(* IEC 61131-3 sources: daoli-st-library/DL_Process (part 59) *)

(* ---- FB_DL_WaferThermalBudgetAccum.st ---- *)
(*==============================================================================
 * 组件名称 (Component)  : FB_DL_WaferThermalBudgetAccum
 * 所属子库 (Sublibrary) : DL_Process
 * 归属目录 (Directory)  : C:\Library\DL_Process
 * 当前版本 (Version)    : 1.0.1
 * 分类/来源标签         : 功能块（FUNCTION_BLOCK）· 半导体热预算 · Arrhenius 积分
 *                         industry-pool / semiconductor / thermal-budget
 * 兼容性   (Platform)   : CODESYS 3.5 / TwinCAT 3 / 汇川 InoProShop / 施耐德
 *                         Machine Expert；仅用 Standard.library 的 TON / EXP / ABS
 * 溯源声明 (Provenance) : 道莅自研 clean-room——只借公开规范条款与工程惯例，零代码行复制。
 * 功能一句话 (Summary)  : 晶圆热预算累计：温度对时间的 Arrhenius 加权积分
 *                         （归一到参考温度等效秒），超工艺窗口锁存告警。
 *
 * 量纲链（R25 P2 模板）：
 *   输入 fWaferTempC [degC] → 开尔文 T [K] = fWaferTempC + 273.15
 *   权重 w [无量纲] = EXP(fEaOverK × (1/fTRefK − 1/T))，参考温度处 w 恒为 1
 *   预算 fBudgetEqS [s@fTRefC] = Σ(w × Δt)，Δt 由采样节拍定时器导出 [s]
 *   判据 fBudgetEqS 与 fBudgetLimit [s@fTRefC] 同量纲直接比较
 *
 * 功能描述 (Function)   : 三态状态机：空闲/累计/超限锁存。工艺进行中按节拍
 *                         采样温度，每拍把 w × 节拍秒累入预算；温度非物理
 *                         （≤ −273.15 degC 或非有限）报故障冻结累计；预算超
 *                         上限转入超限相锁存告警（故障级 3025），仅复位指令
 *                         可解除（可达解除路径）；复位以信息级 3023 告知。
 * 与既有件边界 (Boundary): 本件只做预算累计与超限告警，不控温；温控归
 *                         工艺温控环，本件是良率保护层。
 * 码位说明 (Codes)      : 信息 16#0006_3023 预算复位执行，锁存告警解除
 *                         故障 16#0006_3024 温度非物理域（≤ −273.15 degC 或非有限）
 *                         故障 16#0006_3025 热预算超工艺窗口，已锁存告警
 *                         段 16#06_0_23~27 首槽信息级、次槽起故障级。
 * 依赖说明 (Depends)    : 无 DL_ 内部依赖；仅 Standard.library 的 TON / EXP。
 * 红线自检 (Redline)    : 零全局依赖 ｜ 零 VAR_EXTERNAL ｜ 零 %I/%Q ｜ 纯 IEC 标准库
 *                         NaN/Inf 精确判据拦截 ｜ 浮点比较带 fEps 容差
 *                         ENUM 配 CASE 且 ELSE 兜底 ｜ TON 每周期无条件刷新
 *                         全变量双语同行注释 ｜ 量纲链头注释齐备（R25 P2）
 * 修订历史 (Revision)   : 2026-11-18  v1.0.0  首版入库（R32 · 批 4）
 *                        2026-11-18  v1.0.1  R33 返修：温度恢复清 3024；复位沿提前段 1 全局；采样节拍正域闸（≤0 置 3024 跳过累计）
 *============================================================================*)

FUNCTION_BLOCK FB_DL_WaferThermalBudgetAccum
VAR_INPUT
    bRun         : BOOL;                // 累计使能 / Enable
    bInProcess   : BOOL;                // 工艺进行中 [事件]，真才累计 / Process active flag
    fWaferTempC  : LREAL;               // 晶圆温度 [degC] / Wafer temperature
    fTRefC       : LREAL := 200.0;      // 参考温度 [degC]，等效秒归一基准 / Reference temperature
    fEaOverK     : LREAL := 8000.0;     // 活化能除气体常数 [K]，Arrhenius 斜率 / Ea over k in kelvin
    tSample      : TIME  := T#1S;       // 采样节拍 [s] / Sampling pace period
    fBudgetLimit : LREAL := 3600.0;     // 预算上限 [s@fTRefC] / Budget limit in reference seconds
    bReset       : BOOL;                // 复位指令 [事件]，沿触发清预算与锁存 / Reset command, edge triggered
    fEps         : LREAL := 1.0E-6;     // 浮点判零容差 [实数域] / Floating zero tolerance
END_VAR
VAR_OUTPUT
    ePhase    : (ePhaseIdle := 0, ePhaseAccum := 1, ePhaseExceeded := 2);    // 相枚举输出 / Phase output enum
    fBudgetEqS: LREAL;                  // 等效参考秒累计 [s@fTRefC] / Accumulated budget
    fWeightNow: LREAL;                  // 当前权重 [无量纲] / Current Arrhenius weight
    bExceeded : BOOL;                   // 超限锁存告警 / Latched over-limit alarm
    bError    : BOOL;                   // 故障标志，与故障码配对 / Fault flag paired with codes
    uErrorId  : UDINT;                  // 事件码，0 表示无事件 / Event code, zero means none
END_VAR
VAR
    _eState  : (eStIdle := 0, eStAccum := 1, eStExceeded := 2);  // 内部状态机 / Internal state machine
    tonPace  : TON;     // 采样节拍定时器 [s]，每拍无条件刷新 / Sampling pace timer
    rTrigRst : R_TRIG;  // 复位上升沿检测，每拍无条件刷新 / Reset edge detection
    fTK      : LREAL;   // 开尔文温度 [K] / Kelvin temperature
    fTRefK   : LREAL;   // 参考开尔文 [K] / Reference in kelvin
    fDeltaS  : LREAL;   // 本拍等效秒增量 [s@fTRefC] / Budget increment this scan
    bTempOk  : BOOL;    // 温度有效标志 / Temperature validity flag
    fPaceS   : LREAL;   // 节拍秒值 [s]，一次导出 / Pace seconds, derived once
    uCode    : UDINT;   // 码位暂存，出口单点写入 [码] / Code staging
    bTempOkPrev : BOOL; // 上拍温度有效快照，恢复沿判据 / Previous validity snapshot
    bPaceOk  : BOOL;    // 采样节拍正域闸标志（tSample > 0）/ Positive pace domain gate
END_VAR
VAR CONSTANT
    DL_WTA_ABS0 : LREAL := 273.15;      // 绝对零度 [degC] / Absolute zero in celsius
    DL_WTA_MS2S : LREAL := 1000.0;      // 毫秒到秒系数 [ms/s] / Milliseconds per second
END_VAR

(* 段 1｜定时器与边沿无条件刷新 + 全局复位 + 节拍正域闸（R33 返修：复位沿提前到全局，不再只挂 eStExceeded）
 *      Timers and edges refreshed unconditionally, global reset edge, positive pace domain gate *)
tonPace(IN := NOT tonPace.Q, PT := tSample);    // 节拍自复位振荡（红线 7，Q 每节拍单拍脉冲）/ Self-reset pace
rTrigRst(CLK := bReset);                        // 复位沿检测 / Reset edge detection
IF fPaceS < 0.0001 THEN
    fPaceS := DINT_TO_LREAL(TIME_TO_DINT(tSample)) / DL_WTA_MS2S;   // 节拍秒值一次导出 / Derive pace once
END_IF
bPaceOk := (tSample > T#0S) AND (fPaceS > fEps); // 节拍正域闸：≤0 时置 3024 并跳过累计 / Positive pace gate
IF rTrigRst.Q THEN
    (* 全局复位：预算清零、锁存解除、回空闲，任何相均可达 / Global reset reachable from any phase *)
    fBudgetEqS := 0.0;          // 预算清零 / Clear the budget
    bExceeded := FALSE;         // 解除锁存 / Release the latch
    uCode := 16#0006_3023;      // 信息级：复位执行 / Info: reset executed
    _eState := eStIdle;         // 拍 N+1 回空闲重部署 / To idle for redeploy
END_IF

(* 段 2｜温度有效性（NaN 自反、Inf 上限、绝对零物理域）/ Temperature validity *)
fTK := fWaferTempC + DL_WTA_ABS0;               // 摄氏转开尔文 / Celsius to kelvin
fTRefK := fTRefC + DL_WTA_ABS0;                 // 参考转开尔文 / Reference to kelvin
bTempOk := (fWaferTempC = fWaferTempC)          // NaN 自反判据 / NaN reflexivity
           AND (ABS(fWaferTempC) < 1.0E308)     // Inf 上限判据 / Inf limit
           AND (fWaferTempC > -DL_WTA_ABS0)     // 绝对零物理域 / Above absolute zero
           AND (fTRefK > fEps);                 // 参考温度防零除 / Reference above zero
IF bTempOk AND (NOT bTempOkPrev) AND (uCode = 16#0006_3024) THEN
    uCode := 16#0000_0000;          // 温度恢复沿清 3024（复位可达，不动 3025 锁存）/ Recovery clears 3024
END_IF
bTempOkPrev := bTempOk;             // 有效标志快照 / Validity snapshot

(* 段 3｜状态机主分派（ENUM 配 CASE，ELSE 兜底）/ State dispatch with ELSE interception *)
CASE _eState OF

    eStIdle:
        (* 本拍行为：预算保持；使能且数据有效拍 N+1 转累计 / Hold; arm when valid *)
        bExceeded := FALSE;             // 空闲无告警 / No alarm in idle
        IF bRun AND bTempOk AND (NOT bInProcess) THEN
            fBudgetEqS := 0.0;          // 进累计前清预算 / Clear before accumulating
        END_IF
        IF bRun AND bTempOk THEN
            _eState := eStAccum;        // 拍 N 空闲相满足，拍 N+1 转累计 / To accumulating next scan
        END_IF
        IF NOT bTempOk THEN
            uCode := 16#0006_3024;      // 故障级：温度非物理域 / Fault: non-physical temperature
        END_IF

    eStAccum:
        (* 本拍行为：工艺进行中按节拍累加 Arrhenius 权重秒 / Accumulate weighted seconds *)
        IF NOT bRun THEN
            _eState := eStIdle;         // 拍 N+1 回空闲 / To idle next scan
        ELSIF NOT bTempOk THEN
            uCode := 16#0006_3024;      // 故障级：温度非物理域，累计冻结 / Fault: freeze
            bTempOk := FALSE;
        ELSE
            fWeightNow := EXP(fEaOverK * (1.0 / fTRefK - 1.0 / fTK));   // Arrhenius 权重 / Arrhenius weight
            IF bInProcess AND tonPace.Q AND bPaceOk THEN
                fDeltaS := fWeightNow * fPaceS;     // 本拍等效秒增量 / Increment in reference seconds
                fBudgetEqS := fBudgetEqS + fDeltaS; // 预算累加 / Accumulate the budget
            END_IF
            IF NOT bPaceOk THEN
                uCode := 16#0006_3024;  // 节拍非正域（tSample ≤ 0）：置码并跳过累计，禁止静默 / Non-positive pace: code and skip
            END_IF
            IF fBudgetEqS > fBudgetLimit THEN
                _eState := eStExceeded; // 拍 N+1 转超限锁存 / To exceeded next scan
                bExceeded := TRUE;      // 超限告警锁存 / Latch the alarm
                uCode := 16#0006_3025;  // 故障级：预算超限 / Fault: budget exceeded
            END_IF
        END_IF

    eStExceeded:
        (* 本拍行为：停止累计保持告警；解除路径已提前至段 1 全局复位沿（R33 返修）
         * Stop accumulating, keep the alarm; clear path is the global reset edge in segment 1 *)
        bExceeded := TRUE;              // 锁存回放，防止中途被旁路覆盖 / Latch replay
        uCode := 16#0006_3025;          // 故障级回放 / Fault replay

ELSE
    _eState := eStIdle;                 // 非法状态拦截回空闲 / Illegal state to idle
    uCode := 16#0006_3024;              // 故障：状态越界 / Fault: state out of range
END_CASE

(* 段 4｜出口装配 / Exit assembly *)
ePhase := ePhaseIdle;                   // 相映射刷新 / Refresh the phase mapping
IF _eState = eStAccum THEN
    ePhase := ePhaseAccum;
ELSIF _eState = eStExceeded THEN
    ePhase := ePhaseExceeded;
END_IF
bError := (uCode >= 16#0006_3024) AND (uCode <= 16#0006_3025);  // 故障级码带判定 / Fault band check
uErrorId := uCode;                      // 码位单点写入 / Single write point
END_FUNCTION_BLOCK

(* ---- FB_DL_WaterChlorineDoseTrim.st ---- *)
(*
  道莅工业代码库 | DL_Process | FB_DL_WaterChlorineDoseTrim
  版本: 1.0.0 | 日期: 2026-11-23 | 轮次: R75
  开源溯源: self-cleanroom（无外部来源；绿区水处理语义域延伸，零代码行复制）
  功能: 余氯-浊度双参数加药量 trim 控制——以余氯偏差比例 trim 出口加药量设定，
        浊度超高经延时进护栏态（trim 只允许下调禁上调），剂量上限闸（±fTrimLim），
        流量折算加药流量出口（L/h）。
  兼容性: CODESYS 3.5 / TwinCAT 3 / 汇川 InoProShop；仅依赖标准 TON / R_TRIG / LIMIT，零厂商私有库
  接口: 输入余氯实测/设定、浊度实测/上限、基准加药量、trim 增益与幅值限、
        处理流量、周期、冻结、复位；输出 fDoseRate [mg/L]/fTrimOut [mg/L]/
        fDoseFlow [L/h]/bTurbGuard/eState/eCause/bError/nErrId。
  码表: 16#0005_03B9 故障级：传感器非有限（余氯/浊度 NaN，锁存至复位沿，剂量保持最后有效值）
        16#0005_04E0 信息级：处理流量近零（fDoseFlow 出口钳零，加药量出口不受影响）
        码段说明：0005 段故障子带 03xx / 信息子带 04xx，槽位经全库实扫空闲。
  边界: ① trim 幅值闸：LIMIT(±fTrimLim)，护栏态下 trim := MIN(trim, 0)（只降不升）；
        ② 护栏态退出条件 ≥ 2 条：浊度回落前置消失，或使能撤/复位事件；
        ③ 传感器 NaN 故障锁存期间剂量保持锁存量（不随坏值波动）；
        ④ fDoseFlow = fDoseRate·fFlowAct/1000，除法无（乘法），流量比换算在出口
        判 fFlowAct > EPS 否则钳零并置信息码；
        ⑤ TON/R_TRIG 段 0 无条件周期刷新；⑥ 零全局耦合。
  邻件比对: DosingPumpCalib/BatchDosingControl（标定/批量加药 vs 本件余氯连续 trim）。
  修订历史: 2026-11-23 v1.0.0 R75 首版（复杂件批 B2 · C07）
*)

TYPE E_DL_WctState :
(
    eIdle     := 0,   // 待机（出口保持） | Idle, outlet held
    eTrim     := 10,  // 正常 trim 运行 | Normal trim run
    eTurbHold := 20,  // 浊度护栏（trim 禁上调） | Turbidity guard, trim down only
    eFault    := 90   // 故障锁存相 | Fault latch phase
);
END_TYPE

TYPE E_DL_WctCause :
(
    eNone          := 0,  // 无故障 | No cause
    eCfgIllegal    := 1,  // 组态非法 | Illegal configuration
    eSensNonFinite := 2   // 传感器非有限 | Sensor non-finite
);
END_TYPE

FUNCTION_BLOCK FB_DL_WaterChlorineDoseTrim
VAR_INPUT
    bAutoEn   : BOOL := FALSE;    // 自动 trim 使能 [-] | Auto trim enable
    fClResAct : REAL := 0.0;      // 余氯实测 [mg/L] | Chlorine residual actual
    fClResSp  : REAL := 0.8;      // 余氯设定，域 > 0 [mg/L] | Chlorine residual setpoint
    fTurbAct  : REAL := 0.0;      // 浊度实测 [NTU] | Turbidity actual
    fTurbMax  : REAL := 1.0;      // 浊度护栏上限，域 > 0 [NTU] | Turbidity guard limit
    fDoseBase : REAL := 1.2;      // 基准加药量，域 >= 0 [mg/L] | Base dose
    fKpTrim   : REAL := 1.0;      // trim 比例增益，域 >= 0 [mg/L per mg/L] | Trim proportional gain
    fTrimLim  : REAL := 0.5;      // trim 幅值限（±对称），域 >= 0 [mg/L] | Trim magnitude limit
    fFlowAct  : REAL := 0.0;      // 处理流量 [m3/h] | Treated flow actual
    fDtSec    : REAL := 0.1;      // 调节周期（护栏去抖基准），域 (0, 1] [s] | Trim cycle time
    tTurbHold : TIME := T#10S;    // 浊度超高确认延时，域 > T#0S | Turbidity confirm delay
    bFreeze   : BOOL := FALSE;    // trim 冻结（电平，剂量回基准）[-] | Trim freeze level
    bReset    : BOOL := FALSE;    // 复位命令，上升沿清故障 [-] | Reset command, rising edge
END_VAR
VAR_OUTPUT
    fDoseRate  : REAL;            // 出口加药量设定 [mg/L] | Dose rate outlet
    fTrimOut   : REAL;            // trim 分量出口 [mg/L] | Trim component outlet
    fDoseFlow  : REAL;            // 折算加药流量出口 [L/h] | Dosing flow outlet
    bTurbGuard : BOOL;            // 浊度护栏激活态 [-] | Turbidity guard active
    eState     : E_DL_WctState;   // 状态出口 | State outlet
    eCause     : E_DL_WctCause;   // 故障成因出口 | Fault cause outlet
    bError     : BOOL;            // 故障锁存标志 [-] | Fault latch flag
    nErrId     : UDINT;           // 事件码，0 = 无事件 | Event code, 0 = none
END_VAR
VAR
    _eState   : E_DL_WctState := E_DL_WctState.eIdle;   // 内部状态（CASE 唯一写入目标） | Internal state
    _eCause   : E_DL_WctCause := E_DL_WctCause.eNone;   // 成因锁存 | Latched cause
    _bFault   : BOOL;             // 故障锁存位 | Fault latch bit
    _fDoseRate: REAL := 0.0;      // 剂量锁存量 [mg/L]（故障保持载体） | Dose rate latch
    _fTrimOut : REAL := 0.0;      // trim 锁存量 [mg/L]（故障保持载体） | Trim latch
    _bCfgBad  : BOOL;             // 组态非法当拍量 [-] | Illegal configuration
    _bSensBad : BOOL;             // 传感器非有限当拍量 [-] | Sensor non-finite this scan
    _bTurbHi  : BOOL;             // 浊度超高当拍量 [-] | Turbidity high this scan
    _bFlowLo  : BOOL;             // 流量近零当拍量 [-] | Flow near zero this scan
    _uInfo    : UDINT;            // 信息码每拍重算 | Info code per scan
    fErr      : REAL;             // 余氯偏差当拍量 [mg/L] | Residual error this scan
    fTrimCalc : REAL;             // 本拍 trim 计算量 [mg/L] | Trim calculated this scan
    rtReset   : R_TRIG;           // 复位沿实例，段 0 无条件刷新 | Reset edge instance
    tonTurb   : TON;              // 浊度超高确认计时，段 0 无条件刷新 | Turbidity confirm timer
END_VAR
VAR CONSTANT
    DL_WCT_EPS : REAL := 1.0E-6;      // 流量近零判据 [m3/h] | Flow zero threshold
    DL_WCT_ERR : UDINT := 16#0005_03B9;   // 传感器非有限故障码 | Sensor non-finite code
    DL_WCT_IFL : UDINT := 16#0005_04E0;   // 流量近零信息码 | Flow near-zero info code
END_VAR

(* —— 段 0：当拍量派生 + 定时器与沿实例无条件周期刷新（R7 红线） —— *)
_bSensBad := (fClResAct <> fClResAct) OR (fTurbAct <> fTurbAct);            // 传感器 NaN 自反判 / Sensor NaN self-reflex check
_bCfgBad := (fClResSp <= 0.0) OR (fTurbMax <= 0.0) OR (fDoseBase < 0.0)
         OR (fKpTrim < 0.0) OR (fTrimLim < 0.0) OR (fDtSec <= 0.0) OR (fDtSec > 1.0);  // 组态域闸 / Configuration gate
_bTurbHi := (NOT _bSensBad) AND (fTurbAct > fTurbMax);                      // 浊度超高判据（NaN 不判超高） / Turbidity high judgement
_bFlowLo := (fFlowAct <= DL_WCT_EPS) OR (fFlowAct <> fFlowAct);             // 流量近零/非有限判据 / Flow near-zero or non-finite
rtReset(CLK := bReset);                                                     // 复位沿每拍必调 / Reset edge every scan
tonTurb(IN := bAutoEn AND _bTurbHi, PT := tTurbHold);                       // 浊度去抖 IN 挂使能 ∧ 超高 / Debounce gated by enable and turbidity

(* —— 段 1：单拍量预清零 —— *)
_uInfo := 16#0000_0000;                                                     // 信息码每拍重算 / Info recomputed per scan
fErr := 0.0;                                                                // 偏差当拍量预清 / Error preset
fTrimCalc := 0.0;                                                           // trim 计算量预清 / Trim calc preset

(* —— 段 2：复位沿 + 组态/传感器域闸 —— *)
IF rtReset.Q AND (NOT _bCfgBad) THEN                                        // 复位沿且组态合法 / Reset with legal config
    _bFault := FALSE;                                                       // 清故障锁存位 / Clear fault latch
    _eCause := E_DL_WctCause.eNone;                                         // 清成因 / Clear cause
    IF _eState = E_DL_WctState.eFault THEN
        _eState := E_DL_WctState.eIdle;                                     // 故障相迁出唯一路径 / Sole fault exit
    END_IF
END_IF
IF _bCfgBad THEN                                                            // 组态域闸 / Configuration gate
    _bFault := TRUE;
    _eCause := E_DL_WctCause.eCfgIllegal;                                   // 归因组态 / Cause: config
END_IF
IF _bSensBad AND (NOT _bFault) THEN                                         // 传感器域闸（组态闸优先归因） / Sensor gate
    _bFault := TRUE;
    _eCause := E_DL_WctCause.eSensNonFinite;                                // 归因传感器 / Cause: sensor
END_IF

(* —— 段 3：trim 计算（限幅 + 护栏只降 + 冻结归零） —— *)
IF bAutoEn AND (NOT _bFault) AND (NOT _bSensBad) THEN
    fErr := fClResSp - fClResAct;                                           // 余氯偏差（正=欠氯需增药）[mg/L] / Residual error
    fTrimCalc := fKpTrim * fErr;                                            // 比例 trim 计算 [mg/L] / Proportional trim
    fTrimCalc := LIMIT(-fTrimLim, fTrimCalc, fTrimLim);                     // 剂量幅值闸（±对称限幅） / Magnitude gate
    IF _bTurbHi THEN
        fTrimCalc := 0.5 * (fTrimCalc + MIN(fTrimCalc, 0.0));               // 护栏半限：向零收敛、只允许下调分量 / Guard: converge toward zero, down-only
    END_IF
    IF bFreeze THEN
        fTrimCalc := 0.0;                                                   // 冻结：trim 归零（剂量回基准） / Freeze: trim zero
    END_IF
    _fTrimOut := fTrimCalc;                                                 // trim 锁存量更新（有效拍才写） / Trim latch updated on valid scans
    _fDoseRate := fDoseBase + _fTrimOut;                                    // 剂量 = 基准 + trim [mg/L] / Dose = base + trim
    IF _fDoseRate < 0.0 THEN
        _fDoseRate := 0.0;                                                  // 剂量非负防御（基准+负 trim 越界） / Dose non-negative defense
    END_IF
END_IF

(* —— 段 4：状态机（ENUM + CASE，ELSE 兜底） —— *)
CASE _eState OF

E_DL_WctState.eIdle:
    IF bAutoEn AND (NOT _bFault) THEN
        _eState := E_DL_WctState.eTrim;                                     // 使能进 trim / Enabled, enter trim
    END_IF

E_DL_WctState.eTrim:
    IF tonTurb.Q THEN
        _eState := E_DL_WctState.eTurbHold;                                 // 浊度超高确认进护栏 / Turbidity confirmed, guard
    ELSIF (NOT bAutoEn) OR _bFault THEN
        _eState := E_DL_WctState.eIdle;                                     // 使能撤或故障回待机 / Disable or fault, idle
    END_IF

E_DL_WctState.eTurbHold:
    IF (NOT _bTurbHi) OR (NOT bAutoEn) THEN
        _eState := E_DL_WctState.eTrim;                                     // 退出双条件：浊度回落（去抖经 tonTurb 重入）或使能撤 / Dual exit conditions
    ELSIF _bFault THEN
        _eState := E_DL_WctState.eIdle;                                     // 故障回待机 / Fault, idle
    END_IF

E_DL_WctState.eFault:
    ;                                                                       // 剂量保持锁存量（故障冻结）/ Dose holds latch, only reset leaves

ELSE
    _bFault := TRUE;                                                        // 非法状态兜底（R6）/ Illegal state fallback
    _eCause := E_DL_WctCause.eCfgIllegal;                                   // 归因归并组态 / Cause folded to config
    _eState := E_DL_WctState.eFault;

END_CASE

(* —— 段 5：故障锁存状态迁移闸 —— *)
IF _bFault AND (_eState <> E_DL_WctState.eFault) THEN
    _eState := E_DL_WctState.eFault;                                        // 锁存即入故障相（剂量冻结在锁存量）/ Latch enters fault phase
END_IF

(* —— 段 6：出口单点映射（名实同源；锁存码回放） —— *)
fDoseRate := _fDoseRate;                                                    // 剂量出口（故障相回放锁存量）[mg/L] / Dose outlet
fTrimOut := _fTrimOut;                                                      // trim 出口 [mg/L] / Trim outlet
IF _bFlowLo OR _bFault THEN
    fDoseFlow := 0.0;                                                       // 流量近零/故障折算出口钳零 [L/h] / Flow outlet clamped zero
    IF _bFlowLo THEN
        _uInfo := DL_WCT_IFL;                                               // 信息级：流量近零 / Info: flow near zero
    END_IF
ELSE
    fDoseFlow := _fDoseRate * fFlowAct * 0.001;                             // 折算加药流量 = 剂量·流量/1000 [L/h] / Dosing flow conversion
END_IF
bTurbGuard := (_eState = E_DL_WctState.eTurbHold);                          // 护栏镜像 / Guard mirror
eState := _eState;                                                          // 状态出口 / State outlet
eCause := _eCause;                                                          // 成因出口 / Cause outlet
bError := _bFault;                                                          // 故障标志同源 / Error flag from latch
IF _bFault THEN
    nErrId := DL_WCT_ERR;                                                   // 故障锁存码回放 / Replay latched fault code
ELSE
    nErrId := _uInfo;                                                       // 信息码 / Info code
END_IF

END_FUNCTION_BLOCK

(* ---- FB_DL_WeighHopperRefillSeq.st ---- *)
(*
  ============================================================
  组件名 : FB_DL_WeighHopperRefillSeq
  分类   : DL_Process
  功能   : 料斗补料顺序控制，开阀快加慢加关阀稳定，含阀超时、稳定超时与人工停止故障
  开源溯源 : internal-design（本轮无外部代码逐行引用）
             参考语义 : 无外部参考
  复杂度 : C2
  版本   : 1.0.0
  ============================================================
*)

TYPE E_DL_HopperState :
(
    eIdle      := 0, // 待机，等待启动命令 idle awaiting the start command
    eValveOpen := 1, // 开阀建流单拍相 the single scan valve opening phase
    eFastFeed  := 2, // 快速加料相 the fast feed phase
    eSlowFeed  := 3, // 慢速加料相 the slow feed phase
    eSettle    := 4, // 关阀后稳定相 the settle phase after the valve closes
    eFault     := 5, // 故障锁存相 the latched fault phase
    eDone      := 6  // 配料完成相 the dosing done phase
);
END_TYPE

FUNCTION_BLOCK FB_DL_WeighHopperRefillSeq
VAR_INPUT
    bStart         : BOOL; // 启动命令 start command
    bStop          : BOOL; // 停止命令 stop command
    rWeight        : REAL; // 料斗实测重量 [kg] measured hopper weight [kg]
    rTargetHigh    : REAL; // 高料位目标 [kg] high level target [kg]
    rTargetLow     : REAL; // 快慢切换点 [kg] fast to slow switching point [kg]
    rSettleBand    : REAL; // 稳定允差带 [kg] settle band [kg]
    tValveTimeout  : TIME; // 加料阀超时窗 [ms] feed valve timeout window
    tSettleTimeout : TIME; // 稳定超时窗 [ms] settle timeout window
END_VAR
VAR_OUTPUT
    bValveOpen : BOOL; // 加料阀开命令 feed valve open command
    bFastFeed  : BOOL; // 快加料命令 fast feed command
    bSlowFeed  : BOOL; // 慢加料命令 slow feed command
    eState     : E_DL_HopperState; // 当前状态 current state
    bDone      : BOOL; // 完成标志，保持到复位沿 done flag held until the reset edge
    nFaultCode : INT; // 故障码 0无 1阀超时 2稳定超时 3人工停止 [码] fault code 0 none, 1 valve, 2 settle, 3 manual stop [code]
END_VAR
VAR
    _eState  : E_DL_HopperState := E_DL_HopperState.eIdle; // 内部状态 internal state
    _bDone   : BOOL := FALSE; // 完成锁存内部量 internal done latch
    _nFault  : INT := 0; // 故障码锁存内部量 latched fault code
    _rBand   : REAL := 0.0; // 钳位后的稳定带 [kg] clamped settle band [kg]
    tonValve : TON; // 加料阀累计超时计时 accumulated valve timeout timer
    tonSettle: TON; // 稳定超时计时 settle timeout timer
    rtStart  : R_TRIG; // 启动命令上升沿 start command rising edge
    rtStop   : R_TRIG; // 停止命令上升沿 stop command rising edge
END_VAR

// 段 0｜定时器与沿实例无条件周期刷新 unconditional cyclic refresh of timers and edges
rtStart(CLK := bStart); // 启动沿刷新 refresh the start edge
rtStop(CLK := bStop); // 停止沿刷新 refresh the stop edge
tonValve(IN := ((_eState = E_DL_HopperState.eValveOpen) OR (_eState = E_DL_HopperState.eFastFeed) OR (_eState = E_DL_HopperState.eSlowFeed)) AND (_nFault = 0), PT := tValveTimeout); // 加料阀累计超时 valve cumulative timeout
tonSettle(IN := (_eState = E_DL_HopperState.eSettle) AND (_nFault = 0), PT := tSettleTimeout); // 稳定超时 settle timeout
// 段 1｜出口预置与输入整形 preset the outputs and reshape the inputs
bValveOpen := FALSE; // 阀命令每拍先关 valve command closed each scan first
bFastFeed := FALSE; // 快加命令每拍先关 fast feed off each scan first
bSlowFeed := FALSE; // 慢加命令每拍先关 slow feed off each scan first
_rBand := rSettleBand; // 取入参稳定带 take the settle band input
IF _rBand < 0.0 THEN
    _rBand := ABS(_rBand); // 负稳定带取幅值 a negative band becomes its magnitude
END_IF
IF (rWeight <> rWeight) OR (rTargetHigh <> rTargetHigh) OR (rTargetLow <> rTargetLow) OR (rSettleBand <> rSettleBand) THEN
    eState := _eState; // 非有限测量或组态拒收，状态保持 refuse a non finite reading or configuration and hold the state
    bDone := _bDone; // 完成标志按锁存量输出 map the latched done flag
    nFaultCode := _nFault; // 故障码按锁存量输出 map the latched fault code
    RETURN; // 早退保护 early return for protection
END_IF
// 段 2｜停止命令优先消化，置于状态机之前 stop command digested ahead of the state machine
IF bStop AND (_eState <> E_DL_HopperState.eFault) THEN
    _nFault := 3; // 人工停止故障码 manual stop fault code
    _eState := E_DL_HopperState.eFault; // 立即迁入故障相 migrate to the fault phase at once
END_IF
// 段 3｜主状态机 main state machine
CASE _eState OF
E_DL_HopperState.eIdle: // 待机 idle
    _bDone := FALSE; // 待机相清完成锁存 clear the done latch while idle
    IF rtStart.Q AND (NOT bStop) THEN
        _eState := E_DL_HopperState.eValveOpen; // 启动沿有效则迁开阀 a valid start edge opens the valve phase
    END_IF
E_DL_HopperState.eValveOpen: // 开阀建流单拍相 single scan valve opening phase
    bValveOpen := TRUE; // 本拍只开阀 this scan only opens the valve
    _eState := E_DL_HopperState.eFastFeed; // 拍 N 进入开阀相，本拍行为只建流不作重量判据，拍 N+1 转出至快加相
E_DL_HopperState.eFastFeed: // 快速加料相 fast feed phase
    bValveOpen := TRUE; // 阀保持开 the valve stays open
    bFastFeed := TRUE; // 快加料输出有效 the fast feed output is active
    IF rWeight >= rTargetHigh THEN
        _eState := E_DL_HopperState.eSettle; // 到高料位关阀转稳定 the high target closes the valve and starts the settle phase
    ELSIF rWeight >= rTargetLow THEN
        _eState := E_DL_HopperState.eSlowFeed; // 到切换点转慢加 the switching point starts the slow feed phase
    END_IF
E_DL_HopperState.eSlowFeed: // 慢速加料相 slow feed phase
    bValveOpen := TRUE; // 阀保持开 the valve stays open
    bSlowFeed := TRUE; // 慢加料输出有效 the slow feed output is active
    IF rWeight >= rTargetHigh THEN
        _eState := E_DL_HopperState.eSettle; // 到高料位关阀转稳定 the high target closes the valve and starts the settle phase
    END_IF
E_DL_HopperState.eSettle: // 关阀后稳定相 settle phase after the valve closes
    IF ABS(rWeight - rTargetHigh) <= _rBand THEN
        _bDone := TRUE; // 稳定带内判完成 a weight inside the band completes the dosing
        _eState := E_DL_HopperState.eDone; // 迁完成相 migrate to the done phase
    ELSIF tonSettle.Q THEN
        _nFault := 2; // 稳定超时故障码 settle timeout fault code
        _eState := E_DL_HopperState.eFault; // 迁故障相 migrate to the fault phase
    END_IF
E_DL_HopperState.eDone: // 配料完成相 dosing done phase
    IF NOT bStart THEN
        _bDone := FALSE; // 启动命令消失清完成锁存 a vanished start command clears the done latch
        _eState := E_DL_HopperState.eIdle; // 回待机 return to idle
    END_IF
E_DL_HopperState.eFault: // 故障锁存相 latched fault phase
    IF rtStop.Q OR (rtStart.Q AND (NOT bStop)) THEN
        _nFault := 0; // 复位清故障码 the reset edge clears the fault code
        _bDone := FALSE; // 复位清完成锁存 the reset edge clears the done latch
        _eState := E_DL_HopperState.eIdle; // 复位回待机 the reset edge returns to idle
    END_IF
ELSE // 非法状态枚举兜底 the illegal state fallback
    _eState := E_DL_HopperState.eIdle; // 非法状态回落待机 an illegal state falls back to idle
END_CASE
// 段 4｜加料阀累计超时看门狗 the accumulated feed valve watchdog
IF tonValve.Q AND ((_eState = E_DL_HopperState.eFastFeed) OR (_eState = E_DL_HopperState.eSlowFeed) OR (_eState = E_DL_HopperState.eValveOpen)) THEN
    _nFault := 1; // 阀超时故障码 valve timeout fault code
    _eState := E_DL_HopperState.eFault; // 迁故障相 migrate to the fault phase
END_IF
// 段 5｜统一出口映射 the unified exit mapping
bDone := _bDone; // 完成标志出口 map the done flag
nFaultCode := _nFault; // 故障码出口 map the fault code
eState := _eState; // 状态出口 map the state
END_FUNCTION_BLOCK

(* ---- FB_DL_WeightCheckReject.st ---- *)
//==============================================================================
// 功能块：FB_DL_WeightCheckReject ｜ 中文名称：动态称重与剔除控制
// 所属子库：DL_Process ｜ 版本：v1.0.0 ｜ 兼容：CODESYS V3.5+ / TwinCAT 3 / 汇川 InoProShop
// 功能描述：包装线动态称重站：滑动窗均值滤波 → 欠重/合格/超重分级 → 剔除指令与
//           完成反馈握手 → 剔除器拒动检测。无料在位时一律不称重也不判定（空秤 0 g
//           会把「无料」判成「欠重」并触发剔除，是本件的核心防错点）。稳定等待以
//           调用方注入的扫描间隔累加计时，与任务周期解耦；剔除反馈窗用 TON 计时。
//           本件不做重量分选配方管理、不驱动称重仪表、不控输送线主传动（停线仅给
//           建议位 bStopLine，最终是否停线由线控层决定）。
// 开源溯源 (Origin)：道莅原创实现（参考 公开工程惯例 分类与参数域）
// 单位表：重量[g] / 剔除反馈窗[s] / 称重稳定等待[ms] / 扫描间隔[ms] / 样本数[个] /
//         计数[件]
// 错误码表：16#0005_0402 信息级（滤波窗有效样本不足 nFilterSamples，本拍不判、不给
//           剔除命令，不置 bError）/ 16#0005_0403 信息级（无料在位，跳过称重并清滤波
//           窗，不置 bError）/ 16#0005_0345 故障级（合格域上下限倒置 fWeightMinG >=
//           fWeightMaxG，置 bError）/ 16#0005_0346 故障级（剔除器拒动：剔除指令发出后
//           反馈窗内无 bRejectFb，置 bError + bRejectFailed + bStopLine 锁存）/
//           16#0005_0347 故障级（输入非有限独立分支显式映射入本槽，且兼作状态机 ELSE
//           非法状态兜底）。非有限与非法状态共用 0347 的反证句：二者在现有输出组合下
//           不可观测出差异——均为 bError+t 全部输出撤（剔除命令撤、bPass 撤、bValid
//           撤），bStopLine 不因非有限而置位，故 §3 未另给独立槽，本件显式复用不越段。
// 状态机：E_DL_WeightRejectState（eIdle=0 待机 / eSettling=10 稳定等待 /
//           eJudging=20 判定 / eRejecting=30 剔除握手 / eFault=99 故障兜底），
//           CASE 含 ELSE 兜底，ELSE 置 0347 且剔除命令与许可全部撤销。
// 边界行为：① bProductPresent := FALSE → 不判定、撤销剔除命令、清滤波窗（防空秤样本
//           污染下一件）+ 信息 0403；② 有效样本 < nFilterSamples → bValid := FALSE +
//           信息 0402，本拍不判且不给剔除命令；③ fWeightMinG >= fWeightMaxG（容差判）
//           → 故障 0345；④ 剔除指令发出后 tRejectWindow 内无反馈 → 故障 0346 +
//           bRejectFailed + bStopLine := TRUE 锁存（漏剔流入下游属安全级，只建议停线
//           不直接停线）；⑤ 非有限（NaN 自反判 + Inf 幅值上限判）→ 独立分支显式置
//           0347，剔除命令撤、许可撤；⑥ 同一件只判一次（bJudged 锁存，料离开才清），
//           防欠重件滞留时反复剔除与反复报拒动；⑦ 失能 → 剔除命令撤 + bPass := FALSE
//           + bValid := FALSE（R72），计数与停线建议锁存保留。
// 修订历史：v1.0.0 2026-11-17 首版（R25 派单 · §4.12）
//==============================================================================
(*------------------------------------------------------------------------------
 * 枚举: E_DL_WeightRejectState（归属 DL_Process，与 FB_DL_WeightCheckReject 同文件）
 *----------------------------------------------------------------------------*)
TYPE E_DL_WeightRejectState :
(
    eIdle      := 0,   // 待机：无料或失能，剔除命令撤 / Idle: no product or disabled, reject command dropped
    eSettling  := 10,  // 稳定等待：料在位但未达 tSettle，不采样 / Settling: product present, sampling not yet allowed
    eJudging   := 20,  // 判定：按滑窗均值分级 / Judging: grading on the sliding-window mean
    eRejecting := 30,  // 剔除握手：命令已发，等反馈 / Rejecting: command issued, waiting for feedback
    eFault     := 99   // 故障兜底：拒动/组态非法/非有限/非法状态 / Fault fallback
);
END_TYPE

(*==============================================================================
 * 功能块: FB_DL_WeightCheckReject
 * 调用约定: 每个扫描周期无条件调用一次；uDeltaTimeMs 必须注入真实任务间隔。
 *============================================================================*)
FUNCTION_BLOCK FB_DL_WeightCheckReject
VAR_INPUT
    fWeightG        : LREAL;                      // 毛重实测 [g] / Gross weight measured [g]
    fWeightMinG     : LREAL;                      // 合格域下限 [g] / Acceptable weight floor [g]
    fWeightMaxG     : LREAL;                      // 合格域上限 [g] / Acceptable weight ceiling [g]
    nFilterSamples  : INT := 5;                   // 滤波窗样本数 [个]，合法域 1~15，域外钳位 / Filter window length [samples], domain 1..15, clamped
    bProductPresent : BOOL;                       // 产品在位（称重台上有料）/ Product present on the weighing platform
    bRejectFb       : BOOL;                       // 剔除完成反馈 / Reject completed feedback
    tRejectWindow   : TIME := T#500MS;            // 剔除反馈窗 [ms]，窗内无反馈判拒动 / Reject feedback window [ms]
    tSettle         : TIME := T#200MS;            // 称重稳定等待 [ms] / Weighing settle time [ms]
    uDeltaTimeMs    : UDINT;                      // 扫描间隔 [ms]，调用方注入，禁系统时间函数 / Scan interval [ms], caller-injected
    bEnable         : BOOL;                       // 总使能 / Master enable
    bReset          : BOOL;                       // 复位，上升沿清拒动锁存、停线建议与计数 / Reset, rising edge clears the reject-failure latch, stop hint and counters
END_VAR
VAR_OUTPUT
    fWeightFilteredG : LREAL;                     // 滑窗均值滤波重量 [g] / Sliding-window mean weight [g]
    bPass           : BOOL;                       // 合格判定（仅本件判过且合格时为 TRUE）/ Pass verdict, TRUE only when judged and within limits
    bRejectCmd      : BOOL;                       // 剔除指令（脉宽 ≥ 反馈窗，命令语义）/ Reject command, held for the feedback window
    nUnderCount     : UDINT;                      // 欠重计数 [件]，饱和 / Underweight counter [pcs], saturating
    nOverCount      : UDINT;                      // 超重计数 [件]，饱和 / Overweight counter [pcs], saturating
    nRejectCount    : UDINT;                      // 剔除指令计数 [件]，饱和（按指令发出口径）/ Reject command counter [pcs], saturating
    bRejectFailed   : BOOL;                       // 剔除器拒动标志（锁存至 bReset）/ Rejector refusal flag, latched until reset
    bNoProduct      : BOOL;                       // 无料在位标志（信息 0403 的出口）/ No-product flag, outlet of info 0403
    bStopLine       : BOOL;                       // 停线建议（只建议不执行，锁存至 bReset）/ Stop-line recommendation only, latched until reset
    eErr            : UDINT;                      // 错误码，0 = 无错，码位 16#0005_0402 起信息级、16#0005_0345 起故障级（分带见错误码表） / Error code, 0 = no error, band info/fault per the code table
    bError          : BOOL;                       // 故障级标志，仅故障级错误置位 / Fault-class flag, set only on fault-level codes
    bValid          : BOOL;                       // 重量结论可用标志，样本不足/失能/故障闸显式 FALSE / Verdict usable flag, explicit FALSE on insufficient samples, disable and fault gates
    eState          : E_DL_WeightRejectState;     // 主状态机当前状态 / Current state of the main state machine
END_VAR
VAR
    fbReset         : R_TRIG;                     // 复位上升沿检测实例 / Reset rising edge detector
    fbTonReject     : TON;                        // 剔除反馈窗定时器实例 / Reject feedback window timer
    afWindow        : ARRAY[0..14] OF LREAL;      // 滑窗样本缓冲 [g]，定长 15 / Sliding-window sample buffer [g], fixed length 15
    nWinIdx         : INT;                        // 滑窗写指针 [—] / Sliding-window write index
    nWinCnt         : INT;                        // 滑窗内有效样本数 [个] / Valid sample count in the window
    nSamplesEff     : INT;                        // 钳位后的滤波窗长度 [个] / Clamped filter length [samples]
    nLoop           : INT;                        // 清零循环索引 [—] / Clearing loop index
    nSampUse        : INT;                        // 本拍参与均值的样本数 [个] / Samples used by the mean this scan
    uSettleAccMs    : UDINT;                      // 稳定等待累计 [ms]，按注入间隔累加 / Settle accumulator [ms], by injected interval
    uSettleMs       : UDINT;                      // 稳定等待目标值 [ms] / Settle target [ms]
    uDtEff          : UDINT;                      // 钳位后的扫描间隔 [ms] / Clamped scan interval [ms]
    uCntMax         : UDINT;                      // 计数器饱和上限 [件] / Counter saturation ceiling [pcs]
    fSumG           : LREAL;                      // 窗口样本求和 [g] / Window sample sum [g]
    bSampleNow      : BOOL;                       // 本拍允许采样 / Sampling allowed this scan
    bSettled        : BOOL;                       // 稳定等待已满足 / Settle time satisfied
    bJudged         : BOOL;                       // 同一件已判定锁存 / One verdict per product latched
    bUnder          : BOOL;                       // 本件欠重判定 / Underweight verdict of this product
    bOver           : BOOL;                       // 本件超重判定 / Overweight verdict of this product
    bRejectAct      : BOOL;                       // 剔除动作进行中（内部）/ Reject action in progress, internal
    bNonFin         : BOOL;                       // 非有限判定中间标志 / Non-finite detection intermediate flag
    bFirstScan      : BOOL := TRUE;               // 上电首拍标志 / First-scan flag
END_VAR
VAR CONSTANT
    DL_WCR_CODE_INFO_1 : UDINT := 16#0005_0402;   // 信息级槽 1（有效样本不足，本拍不判） / info slot 1
    DL_WCR_CODE_INFO_2 : UDINT := 16#0005_0403;   // 信息级槽 2（无料在位跳过称重） / info slot 2
    DL_WCR_CODE_FLT_1  : UDINT := 16#0005_0345;   // 故障级槽 1（合格域上下限倒置） / fault slot 1
    DL_WCR_CODE_FLT_2  : UDINT := 16#0005_0346;   // 故障级槽 2（剔除器拒动） / fault slot 2
    DL_WCR_CODE_FLT_3  : UDINT := 16#0005_0347;   // 故障级槽 3（输入非有限/非法状态兜底） / fault slot 3
    DL_WCR_WIN_MAX     : INT := 15;               // 滤波窗定长上限 [个] / Fixed filter window width [samples]
    DL_WCR_WIN_MIN     : INT := 1;                // 滤波窗下限 [个] / Filter window floor [samples]
    DL_WCR_CNT_MAX     : UDINT := 16#FFFF_FFFE;   // 计数器饱和值 [件] / Counter saturation [pcs]
    DL_WCR_DT_MIN_MS   : UDINT := 1;              // 扫描间隔下限 [ms]，防死等 / Scan interval floor [ms], prevents a dead wait
    DL_WCR_ZERO        : LREAL := 0.0;            // 零值常量，避免裸字面量 [—] / Zero constant, avoids a bare literal
    DL_WCR_TOL         : LREAL := 1.0E-6;         // 浮点比较容差 [—] / Float comparison tolerance
    DL_WCR_INF         : LREAL := 1.7976931348623157E308; // LREAL 幅值上限，Inf 判据 / LREAL magnitude ceiling
    DL_WCR_U32_MAX     : UDINT := 16#FFFF_FFFE;   // 毫秒累加饱和上限 [ms] / Millisecond accumulator saturation [ms]
END_VAR

(*------------------------------------------------------------------------------
 * 段 1｜无条件刷新区（红线 5）：复位沿与剔除窗定时器在任何分支之外周期调用。
 *       定时器 IN 取上拍动作状态（单拍滞后对 ≥500 ms 窗无影响），
 *       保证待机/故障/各分支下计时链永不断流
 *----------------------------------------------------------------------------*)
fbReset(CLK := bReset);                            // 复位沿检测无条件刷新 / reset edge refreshed unconditionally
fbTonReject(IN := bRejectAct AND (NOT bRejectFb),  // 动作中且未收到反馈则计时 / timing while active without feedback
            PT := tRejectWindow);                  // 反馈窗长度 [ms] / feedback window length

(*------------------------------------------------------------------------------
 * 段 2｜复位沿处理（改写置于沿后，防吞沿 R39）
 *----------------------------------------------------------------------------*)
IF fbReset.Q THEN
    eState := E_DL_WeightRejectState.eIdle;
    eErr   := 16#0000_0000;                        // 复位清码 / reset clears the code
    bError := FALSE;                               // 复位清故障 / reset clears the fault
    bRejectFailed := FALSE;                        // 拒动锁存清 / refusal latch cleared
    bStopLine := FALSE;                            // 停线建议清（人工确认后再复位）/ stop hint cleared after manual confirmation
    nUnderCount := 16#0000_0000;                   // 欠重计数清 / underweight counter cleared
    nOverCount := 16#0000_0000;                    // 超重计数清 / overweight counter cleared
    nRejectCount := 16#0000_0000;                  // 剔除计数清 / reject counter cleared
    bRejectAct := FALSE;                           // 动作状态清 / action state cleared
    bJudged := FALSE;                              // 判定锁存清 / verdict latch cleared
    bFirstScan := TRUE;                            // 重新首拍化 / re-initialize first scan
END_IF

(*------------------------------------------------------------------------------
 * 段 3｜非有限输入闸：独立分支显式映射入 0347（头注释给出共用反证句），
 *       剔除命令撤、bPass 撤、bValid 撤；bStopLine 不因非有限置位
 *----------------------------------------------------------------------------*)
bNonFin := (fWeightG <> fWeightG) OR (ABS(fWeightG) >= DL_WCR_INF)
        OR (fWeightMinG <> fWeightMinG) OR (ABS(fWeightMinG) >= DL_WCR_INF)
        OR (fWeightMaxG <> fWeightMaxG) OR (ABS(fWeightMaxG) >= DL_WCR_INF);   // 重量引脚非有限汇总判定 / weight pins non-finite check
IF bNonFin THEN
    eState := E_DL_WeightRejectState.eFault;       // 进故障相 / enter fault state
    eErr   := DL_WCR_CODE_FLT_3;                   // 故障级：输入非有限（显式映射入 0347）/ fault: non-finite input, explicitly mapped onto 0347
    bError := TRUE;                                // 故障级必置 bError（R45 配对）/ fault-class pairs with bError
    bValid := FALSE;                               // 结论不可用 / verdict unusable
    bPass := FALSE;                                // 合格判定撤 / pass verdict dropped
    bRejectCmd := FALSE;                           // 剔除命令撤安全侧 / reject command dropped, safe side
    bRejectAct := FALSE;                           // 动作状态撤 / action state dropped
    fWeightFilteredG := DL_WCR_ZERO;               // 滤波值回零 / filtered value zeroed
    RETURN;
END_IF

(*------------------------------------------------------------------------------
 * 段 4｜组态合法性闸：合格域上下限倒置（容差判，禁浮点判等）
 *----------------------------------------------------------------------------*)
IF (fWeightMinG >= fWeightMaxG - DL_WCR_TOL) THEN
    eState := E_DL_WeightRejectState.eFault;       // 进故障相 / enter fault state
    eErr   := DL_WCR_CODE_FLT_1;                   // 故障级：上下限倒置 / fault: limits inverted
    bError := TRUE;                                // 故障级必置 bError（R45 配对）/ fault-class pairs with bError
    bValid := FALSE;                               // 结论不可用 / verdict unusable
    bPass := FALSE;                                // 合格判定撤 / pass verdict dropped
    bRejectCmd := FALSE;                           // 剔除命令撤安全侧 / reject command dropped, safe side
    bRejectAct := FALSE;                           // 动作状态撤 / action state dropped
    fWeightFilteredG := DL_WCR_ZERO;               // 滤波值回零 / filtered value zeroed
    RETURN;
END_IF

(*------------------------------------------------------------------------------
 * 段 5｜剔除器拒动检测（安全级）：动作中且反馈窗计时到点仍未收到反馈 →
 *       0346 + bRejectFailed + bStopLine 锁存。漏剔会流入下游，故只建议停线
 *       由线控层决策，本件不直接停传动
 *----------------------------------------------------------------------------*)
IF bRejectAct AND fbTonReject.Q AND (NOT bRejectFb) THEN
    bRejectFailed := TRUE;                         // 拒动锁存 / refusal latched
    bStopLine := TRUE;                             // 停线建议锁存（只建议）/ stop-line recommendation latched
    bRejectCmd := FALSE;                           // 剔除命令撤（不再反复打击剔除器）/ command dropped, do not hammer the rejector
    bRejectAct := FALSE;                           // 动作状态撤 / action state dropped
    eState := E_DL_WeightRejectState.eFault;       // 进故障相 / enter fault state
    eErr   := DL_WCR_CODE_FLT_2;                   // 故障级：剔除器拒动 / fault: rejector refused
    bError := TRUE;                                // 故障级必置 bError（R45 配对）/ fault-class pairs with bError
    bValid := FALSE;                               // 结论不可用 / verdict unusable
    RETURN;
END_IF

(*------------------------------------------------------------------------------
 * 段 6｜滤波窗长度钳位与扫描间隔下限（域外按边界钳位，不新占码位：
 *       现有输出组合不可观测出独立信息）
 *----------------------------------------------------------------------------*)
nSamplesEff := nFilterSamples;                     // 先取引脚值 / take the pin value first
IF nSamplesEff < DL_WCR_WIN_MIN THEN
    nSamplesEff := DL_WCR_WIN_MIN;                 // 下限钳位 / clipped to the floor
END_IF
IF nSamplesEff > DL_WCR_WIN_MAX THEN
    nSamplesEff := DL_WCR_WIN_MAX;                 // 上限钳位 / clipped to the ceiling
END_IF
IF uDeltaTimeMs < DL_WCR_DT_MIN_MS THEN
    uDtEff := DL_WCR_DT_MIN_MS;                    // 间隔过小按 1 ms 下限，防稳定等待死等 / floored delta prevents a dead wait
ELSE
    uDtEff := uDeltaTimeMs;                        // 间隔原值 / interval as-is
END_IF
uSettleMs := DINT_TO_UDINT(TIME_TO_DINT(tSettle)); // 稳定等待目标换算 [ms] / settle target in ms

(*------------------------------------------------------------------------------
 * 段 7｜稳定等待累计（按注入间隔，与任务周期解耦）与采样门控
 *----------------------------------------------------------------------------*)
IF bEnable AND bProductPresent THEN
    IF uSettleAccMs < DL_WCR_U32_MAX THEN
        uSettleAccMs := uSettleAccMs + uDtEff;     // 料在位累计稳定时间 [ms] / accumulate settle time while product present
    END_IF
ELSE
    uSettleAccMs := 16#0000_0000;                  // 料离开或失能：稳定计时清零 / product gone or disabled: settle timer cleared
END_IF
bSettled := (uSettleAccMs >= uSettleMs) AND bProductPresent;   // 稳定且料在位 / settled with the product still present
bSampleNow := bEnable AND bProductPresent AND bSettled AND (NOT bJudged);   // 每件在判定前逐拍采样 / sample every scan before the verdict of this product
IF bSampleNow THEN
    afWindow[nWinIdx] := fWeightG;                 // 写入当前样本 [g] / write the current sample
    nWinIdx := nWinIdx + 1;                        // 写指针前移 / advance the write index
    IF nWinIdx >= DL_WCR_WIN_MAX THEN
        nWinIdx := 0;                              // 环形回绕 / ring wrap-around
    END_IF
    IF nWinCnt < DL_WCR_WIN_MAX THEN
        nWinCnt := nWinCnt + 1;                    // 样本计数增（上限 15）/ sample count increments up to 15
    END_IF
END_IF

(*------------------------------------------------------------------------------
 * 段 8｜滑窗均值（只用最近 nSamplesEff 个样本；环形缓冲按逆序回溯取最近样本）
 *----------------------------------------------------------------------------*)
nSampUse := nWinCnt;                               // 先取窗口内有效样本数 / take the valid sample count
IF nSampUse > nSamplesEff THEN
    nSampUse := nSamplesEff;                       // 只用最近 nSamplesEff 个 / use only the newest nSamplesEff samples
END_IF
fSumG := DL_WCR_ZERO;                              // 求和初值 / sum seed
IF nSampUse > 0 THEN
    FOR nLoop := 1 TO nSampUse DO
        fSumG := fSumG + afWindow[(nWinIdx - nLoop + DL_WCR_WIN_MAX * 2) MOD DL_WCR_WIN_MAX];   // 逆序回溯取最近样本 [g] / newest samples in reverse order
    END_FOR
    fWeightFilteredG := fSumG / INT_TO_LREAL(nSampUse);   // 均值（除子已判非零）/ mean, divisor proven non-zero
ELSE
    fWeightFilteredG := DL_WCR_ZERO;               // 无样本时滤波值为 0 / no sample, filtered value zeroed
END_IF

(*------------------------------------------------------------------------------
 * 段 9｜状态机：CASE 含 ELSE 兜底（非法状态 → 0347 + 命令与许可全撤）
 *----------------------------------------------------------------------------*)
CASE eState OF

    E_DL_WeightRejectState.eIdle:
        bRejectCmd := FALSE;                       // 待机剔除命令撤 / reject command dropped in idle
        bRejectAct := FALSE;                       // 动作状态撤 / action state dropped
        bPass := FALSE;                            // 合格判定撤 / pass verdict dropped
        bValid := FALSE;                           // 结论不可用（R72 失能闸）/ verdict unusable on the disable gate
        bNoProduct := NOT bProductPresent;         // 无料标志出口 / no-product flag outlet
        nWinCnt := 0;                              // 无料清窗计数（防空秤污染）/ window count cleared, anti-pollution
        nWinIdx := 0;                              // 写指针复位 / write index reset
        FOR nLoop := 0 TO DL_WCR_WIN_MAX - 1 DO
            afWindow[nLoop] := DL_WCR_ZERO;        // 逐格清零（显式清窗，不留残值）/ explicit per-cell clearing
        END_FOR
        bJudged := FALSE;                          // 判定锁存清（新件重新判）/ verdict latch cleared for the next product
        eErr := 16#0000_0000;                      // 待机无错 / no error in idle
        bError := FALSE;                           // 待机无故障 / no fault in idle
        IF NOT bProductPresent THEN
            eErr := DL_WCR_CODE_INFO_2;            // 信息级：无料在位跳过称重（空秤不出结论）/ info: no product, weighing skipped
        END_IF
        IF bEnable AND bProductPresent THEN
            eState := E_DL_WeightRejectState.eSettling;   // 料在位且使能进稳定等待 / product present and enabled enters settling
        END_IF

    E_DL_WeightRejectState.eSettling:
        bRejectCmd := FALSE;                       // 稳定等待不出剔除 / no reject while settling
        bRejectAct := FALSE;                       // 动作状态撤 / action state dropped
        bPass := FALSE;                            // 未判不出合格 / no pass verdict before judging
        bValid := FALSE;                           // 未判结论不可用 / verdict unusable before judging
        bNoProduct := NOT bProductPresent;         // 无料标志出口 / no-product flag outlet
        eErr := 16#0000_0000;                      // 稳定等待无错 / no error while settling
        bError := FALSE;                           // 稳定等待无故障 / no fault while settling
        IF bEnable AND (NOT bProductPresent) THEN
            eState := E_DL_WeightRejectState.eIdle;   // 料离开回待机（退出条件一）/ product gone, first exit
            eErr := DL_WCR_CODE_INFO_2;            // 信息级：无料在位跳过称重 / info: no product, weighing skipped
        ELSIF bEnable AND bSettled AND (nWinCnt >= nSamplesEff) THEN
            eState := E_DL_WeightRejectState.eJudging;   // 稳定且样本够进判定（退出条件二）/ settled with enough samples, second exit
        END_IF

    E_DL_WeightRejectState.eJudging:
        bError := FALSE;                           // 判定相无故障 / no fault in judging
        bNoProduct := NOT bProductPresent;         // 无料标志出口 / no-product flag outlet
        IF (NOT bProductPresent) THEN
            eState := E_DL_WeightRejectState.eIdle;   // 料离开回待机（退出条件一）/ product gone, first exit
            eErr := DL_WCR_CODE_INFO_2;            // 信息级：无料在位跳过称重 / info: no product, weighing skipped
            bValid := FALSE;                       // 结论不可用 / verdict unusable
            bPass := FALSE;                        // 合格判定撤 / pass verdict dropped
        ELSIF nWinCnt < nSamplesEff THEN
            bValid := FALSE;                       // 样本不足结论不可用（R72）/ insufficient samples, verdict unusable
            bPass := FALSE;                        // 样本不足不判合格 / no pass verdict on insufficient samples
            eErr := DL_WCR_CODE_INFO_1;            // 信息级：有效样本不足，本拍不判 / info: insufficient samples, not judged this scan
            bRejectCmd := FALSE;                   // 样本不足不给剔除命令 / no reject command on insufficient samples
        ELSE
            bValid := TRUE;                        // 样本足够，结论可用 / enough samples, verdict usable
            eErr := 16#0000_0000;                  // 判定相无错 / no error in judging
            IF NOT bJudged THEN
                bUnder := (fWeightFilteredG < fWeightMinG);    // 欠重判据（容差外）/ underweight predicate beyond tolerance
                bOver := (fWeightFilteredG > fWeightMaxG);     // 超重判据（容差外）/ overweight predicate beyond tolerance
                bJudged := TRUE;                   // 本件判定锁存（同件只判一次）/ one verdict per product
                IF bUnder THEN
                    IF nUnderCount < DL_WCR_CNT_MAX THEN
                        nUnderCount := nUnderCount + 1;    // 欠重计数饱和自增 [件] / saturating underweight increment
                    END_IF
                    bPass := FALSE;                // 欠重不合格 / underweight fails
                    bRejectCmd := TRUE;            // 欠重给剔除命令 / reject on underweight
                    bRejectAct := TRUE;            // 动作状态置位（窗计时由此起）/ action state raised, window starts
                    IF nRejectCount < DL_WCR_CNT_MAX THEN
                        nRejectCount := nRejectCount + 1;  // 剔除指令计数 [件] / reject command counter
                    END_IF
                    eState := E_DL_WeightRejectState.eRejecting;   // 进剔除握手相 / enter the reject handshake
                ELSIF bOver THEN
                    IF nOverCount < DL_WCR_CNT_MAX THEN
                        nOverCount := nOverCount + 1;      // 超重计数饱和自增 [件] / saturating overweight increment
                    END_IF
                    bPass := FALSE;                // 超重不合格 / overweight fails
                    bRejectCmd := TRUE;            // 超重给剔除命令 / reject on overweight
                    bRejectAct := TRUE;            // 动作状态置位 / action state raised
                    IF nRejectCount < DL_WCR_CNT_MAX THEN
                        nRejectCount := nRejectCount + 1;  // 剔除指令计数 [件] / reject command counter
                    END_IF
                    eState := E_DL_WeightRejectState.eRejecting;   // 进剔除握手相 / enter the reject handshake
                ELSE
                    bPass := TRUE;                 // 合格放行 / pass and release
                    bRejectCmd := FALSE;           // 合格不剔除 / no reject on pass
                    bRejectAct := FALSE;           // 动作状态撤 / action state dropped
                    eState := E_DL_WeightRejectState.eJudging;     // 留在判定相等料离开 / stay in judging until the product leaves
                END_IF
            ELSE
                bPass := (NOT bUnder) AND (NOT bOver);   // 已判件结论保持 / verdict held for an already-judged product
                IF bUnder OR bOver THEN
                    eState := E_DL_WeightRejectState.eRejecting;   // 不合格件回到握手相等反馈 / unqualified product returns to the handshake
                END_IF
            END_IF
        END_IF

    E_DL_WeightRejectState.eRejecting:
        bValid := TRUE;                            // 结论可用（已判）/ verdict usable, already judged
        bPass := FALSE;                            // 剔除件不合格 / rejected product fails
        bError := FALSE;                           // 握手相无故障（拒动已由段 5 早期判定）/ no fault here, refusal handled earlier
        bRejectCmd := TRUE;                        // 剔除命令保持（脉宽 ≥ 反馈窗）/ command held for at least the feedback window
        bRejectAct := TRUE;                        // 动作状态保持 / action state held
        eErr := 16#0000_0000;                      // 握手相无错 / no error in the handshake
        IF NOT bProductPresent THEN
            bRejectCmd := FALSE;                   // 料已离开：命令撤（退出条件一）/ product gone, first exit
            bRejectAct := FALSE;                   // 动作状态撤 / action state dropped
            eState := E_DL_WeightRejectState.eIdle;   // 回待机 / back to idle
            eErr := DL_WCR_CODE_INFO_2;            // 信息级：无料在位 / info: no product present
        ELSIF bRejectFb THEN
            bRejectCmd := FALSE;                   // 收到反馈：命令撤（退出条件二）/ feedback received, second exit
            bRejectAct := FALSE;                   // 动作状态撤 / action state dropped
            eState := E_DL_WeightRejectState.eJudging;     // 回到判定相等料离开 / back to judging until the product leaves
        END_IF

    E_DL_WeightRejectState.eFault:
        bValid := FALSE;                           // 故障闸显式不可用（R72）/ explicit FALSE on the fault gate
        bPass := FALSE;                            // 合格判定撤 / pass verdict dropped
        bRejectCmd := FALSE;                       // 剔除命令撤安全侧 / reject command dropped, safe side
        bRejectAct := FALSE;                       // 动作状态撤 / action state dropped
        bError := TRUE;                            // 故障级必置 bError（R45 配对）/ fault-class pairs with bError
        IF eErr = 16#0000_0000 THEN
            eErr := DL_WCR_CODE_FLT_3;             // 入口无码时按非法状态兜底（R45：bError 必须有对应码）/ illegal-state fallback so bError always maps to a code
        END_IF
        IF bEnable AND bProductPresent AND (NOT bRejectFailed) THEN
            eState := E_DL_WeightRejectState.eSettling;   // 拒动锁存未清则不得自动恢复；其余条件齐备回稳定等待 / refuse auto-recovery until the latch is cleared
            bJudged := FALSE;                      // 重新判定 / re-judge from scratch
        END_IF

    ELSE
        eState := E_DL_WeightRejectState.eFault;   // 非法状态兜底 / illegal-state fallback
        eErr := DL_WCR_CODE_FLT_3;                 // 故障级兜底：非法状态 / fault fallback: illegal state
        bError := TRUE;                            // 故障级必置 bError（R45 配对）/ fault-class pairs with bError
        bValid := FALSE;                           // 结论不可用 / verdict unusable
        bPass := FALSE;                            // 合格判定撤 / pass verdict dropped
        bRejectCmd := FALSE;                       // 剔除命令撤安全侧 / reject command dropped, safe side
        bRejectAct := FALSE;                       // 动作状态撤 / action state dropped
        fWeightFilteredG := DL_WCR_ZERO;           // 滤波值回零 / filtered value zeroed

END_CASE
END_FUNCTION_BLOCK

(* ---- FB_DL_WeightClassifySort.st ---- *)
// =====================================================================
// FB_DL_WeightClassifySort.st
// 重量四档分级剔除（复用库内判档律 + 剔除口放行 + 档位计数）
// Weight 4-band classification with reject gate and band counters
// 所属子库: DL_Process    版本: v1.0.1    兼容: CODESYS V3.5+ / TwinCAT 3 / 汇川 InoProShop
// 码位: 16#0005_0476 ~ 16#0005_047A (本件独占 5 槽, 勿复用)
// 溯源: 道莅 clean-room 防御性实现
//       来源组标签: packaging, weight-sorting, classification, reject
// 枚举属主: E_DL_WeightClass —— 本文件为全库唯一属主, 其他件只引用不重声明
// 修改记录: R30 初版 (ROUND_PLAN_R30 序 9)
//           v1.0.1 2026-11-23 R75 修复——FC_DL_LimitClassify 调用补
//           uErrorId => uBandErr 显式回执接收（R73 零回执挂账点修），判档件
//           回执非零时按非法档安全侧分流，主判档逻辑零改动
// 分层声明: 判档律消费 DL_Base 的 FC_DL_LimitClassify（四阈值五档, 返回
//           E_DL_LimitBand）, 本件不重写分级律, 只做判档→剔除口→计数编排;
//           区间归属沿用判档件闭区间口径（等于阈值归更严档, 容差判等）
// =====================================================================
// ---------------------------------------------------------------------
// 枚举定义: E_DL_WeightClass (全库唯一属主, 其他件只引用不重声明;
//           R30 序 11 称重剔除秤件引用本枚举)
// ---------------------------------------------------------------------
TYPE E_DL_WeightClass :
(
    eLL,            // 严重欠重档 / Severely underweight band
    eL,             // 欠重档 / Underweight band
    eOK,            // 合格档 / Ok band
    eH,             // 超重档 / Overweight band
    eHH             // 严重超重档 / Severely overweight band
);
END_TYPE

FUNCTION_BLOCK FB_DL_WeightClassifySort
VAR_INPUT
    bPartInZone : BOOL := FALSE;    // 检重区有件信号（分类触发沿）/ Part in check zone, classification trigger
    fWeight_g   : REAL := 0.0;      // 称重值 0~5000 g / Measured weight [g]
    fTh_LL_g    : REAL := 150.0;    // 低低阈值（严重欠重）0~5000 g / Low-low threshold [g]
    fTh_L_g     : REAL := 250.0;    // 低阈值（欠重）0~5000 g / Low threshold [g]
    fTh_H_g     : REAL := 750.0;    // 高阈值（超重）0~5000 g / High threshold [g]
    fTh_HH_g    : REAL := 850.0;    // 高高阈值（严重超重）0~5000 g / High-high threshold [g]
    bRejectArm  : BOOL := FALSE;    // 剔除口布防 / Reject gate armed
END_VAR
VAR_OUTPUT
    eClass      : E_DL_WeightClass := E_DL_WeightClass.eOK;  // 本件判档结果 / Classification result
    bRejectOut  : BOOL := FALSE;    // 剔除口放行脉冲（单拍自清）/ Reject gate pulse, one cycle
    uOkCount    : UDINT := 0;       // 合格计数 / Ok count
    uNgCount    : UDINT := 0;       // 不合格计数（含欠/超重/传感器故障/组态故障安全分流）/ Ng count
    eErr        : UDINT := 16#0005_0476;  // 错误码 / Error code
END_VAR
VAR
    rtrPart     : R_TRIG;           // 有件沿检测, 每拍无条件刷新 / Part edge, refreshed every cycle
    bCfgErr     : BOOL := FALSE;    // 阈值组态非法标记 / Threshold configuration error flag
    eBand       : E_DL_LimitBand := E_DL_LimitBand.eInvalid;  // 判档件返回档 / Band returned by classifier
    bBandInv    : BOOL := FALSE;    // 判档返回非法档标记 / Classifier invalid-band flag
    uBandErr    : UDINT := 0;       // 判档件回执码（v1.0.1 新增接收）/ Classifier receipt code, new in v1.0.1
END_VAR

// ---------------------------------------------------------------------
// 代码位表（本件独占, 勿复用）:
//   16#0005_0476 信息 分级正常（判档完成, OK 或常规 NG 计数）
//   16#0005_0477 故障 阈值组态非法（阈值非有限或越出 0~5000 g 域, 或判档件
//                返回非法档: 阈值序倒置）; 解除式 = 恢复合法单调阈值组态
//   16#0005_0478 故障 重量非有限（传感器故障, NG 侧安全分流, 与超重 NG 区分）,
//                解除式 = 称重值恢复有限且量程内
//   16#0005_0479 信息 超量程（负重为负或超 5000 g, 按 NG 安全分流计数）
//   16#0005_047A 信息 剔除脉冲输出拍（单拍信息, 随剔除口放行同拍发出）
// ---------------------------------------------------------------------

// ---- 有件沿实例无条件刷新 / Unconditional part edge refresh ----
rtrPart(CLK := bPartInZone);

// ---- 阈值组态闸: 四阈值逐一判非有限与量程域（单调性交由判档件校验）
//      Threshold config gate: finite and domain check per threshold ----
bCfgErr := FALSE;                   // 组态标记复位 / Reset config flag
IF (fTh_LL_g <> fTh_LL_g) OR (fTh_LL_g < 0.0) OR (fTh_LL_g > 5000.0) THEN
    bCfgErr := TRUE;                // 低低阈值非法 / Low-low threshold illegal
END_IF
IF (fTh_L_g <> fTh_L_g) OR (fTh_L_g < 0.0) OR (fTh_L_g > 5000.0) THEN
    bCfgErr := TRUE;                // 低阈值非法 / Low threshold illegal
END_IF
IF (fTh_H_g <> fTh_H_g) OR (fTh_H_g < 0.0) OR (fTh_H_g > 5000.0) THEN
    bCfgErr := TRUE;                // 高阈值非法 / High threshold illegal
END_IF
IF (fTh_HH_g <> fTh_HH_g) OR (fTh_HH_g < 0.0) OR (fTh_HH_g > 5000.0) THEN
    bCfgErr := TRUE;                // 高高阈值非法 / High-high threshold illegal
END_IF

// ---- 剔除口缺省收口（单拍脉冲当拍自清）/ Reject pulse default off, self-clearing ----
bRejectOut := FALSE;
bBandInv := FALSE;                  // 非法档标记复位 / Reset invalid-band flag

// ---- 有件沿触发判档编排 / Part edge triggers classification orchestration ----
IF rtrPart.Q THEN
    IF (fWeight_g <> fWeight_g) OR (ABS(fWeight_g) >= 1.0E12) THEN
        // 传感器故障: NG 侧安全分流, 独立故障码 / Sensor fault: NG safe routing, distinct code
        eClass := E_DL_WeightClass.eLL;     // 分流到欠重侧 / Route to underweight side
        bRejectOut := bRejectArm;           // 布防时剔除 / Reject when armed
        uNgCount := uNgCount + 1;           // NG 计数 / Count NG
        eErr := 16#0005_0478;               // 传感器故障码 / Sensor fault code
    ELSIF (fWeight_g < 0.0) OR (fWeight_g > 5000.0) THEN
        // 超量程（含负重为负）: NG 安全分流 / Out of range incl. negative: NG safe routing
        eClass := E_DL_WeightClass.eHH;     // 分流到超重侧 / Route to overweight side
        bRejectOut := bRejectArm;
        uNgCount := uNgCount + 1;
        eErr := 16#0005_0479;               // 超量程信息码 / Over-range info code
    ELSIF bCfgErr THEN
        // 组态故障: 安全侧拒绝分档, 按 NG 分流 / Config fault: safe side, route as NG
        eClass := E_DL_WeightClass.eLL;
        bRejectOut := bRejectArm;
        uNgCount := uNgCount + 1;
        eErr := 16#0005_0477;               // 组态故障码 / Config fault code
    ELSE
        // 判档律消费: 调 DL_Base 判档函数, 闭区间口径 / Consume classifier, closed-interval convention
        eBand := FC_DL_LimitClassify(REAL_TO_LREAL(fWeight_g),
                                     REAL_TO_LREAL(fTh_LL_g),
                                     REAL_TO_LREAL(fTh_L_g),
                                     REAL_TO_LREAL(fTh_H_g),
                                     REAL_TO_LREAL(fTh_HH_g),
                                     uErrorId => uBandErr);   // 回执显式接收（v1.0.1）/ Explicit output receipt
        CASE eBand OF
            E_DL_LimitBand.eLowTripped:     // 低低档 → 严重欠重 / Low-low to severely under
                eClass := E_DL_WeightClass.eLL;
            E_DL_LimitBand.eLowWarn:        // 低档 → 欠重 / Low to under
                eClass := E_DL_WeightClass.eL;
            E_DL_LimitBand.eNormal:         // 正常档 → 合格 / Normal to ok
                eClass := E_DL_WeightClass.eOK;
            E_DL_LimitBand.eUpWarn:         // 高档 → 超重 / High to over
                eClass := E_DL_WeightClass.eH;
            E_DL_LimitBand.eUpTripped:      // 高高档 → 严重超重 / High-high to severely over
                eClass := E_DL_WeightClass.eHH;
            ELSE                            // 非法档兜底: NG 安全侧 / Invalid band fallback: NG safe side
                eClass := E_DL_WeightClass.eLL;
                bBandInv := TRUE;           // 置非法档标记 / Set invalid-band flag
        END_CASE
        IF uBandErr <> 0 THEN               // 判档件回执非零: 按非法档安全侧（v1.0.1 语义接入）/ Classifier receipt nonzero: safe side
            bBandInv := TRUE;               // 置非法档标记 / Set invalid-band flag
        END_IF
        // 档位计数与剔除口放行 / Band counting and reject gate
        IF eClass = E_DL_WeightClass.eOK THEN
            uOkCount := uOkCount + 1;       // 合格计数 / Count ok
        ELSE
            uNgCount := uNgCount + 1;       // 不合格计数 / Count ng
        END_IF
        bRejectOut := bRejectArm AND (eClass <> E_DL_WeightClass.eOK);  // 非 OK 布防剔除 / Reject non-ok when armed
        IF bBandInv THEN
            eErr := 16#0005_0477;           // 判档非法兜底码 / Invalid band code
        ELSE
            eErr := 16#0005_0476;           // 分级正常 / Classification normal
        END_IF
    END_IF
END_IF

END_FUNCTION_BLOCK

(* ---- FB_DL_AerationBlowerCycle.st ---- *)
(*==============================================================================
 * 组件名称 (Component)  : FB_DL_AerationBlowerCycle
 * 所属子库 (Sublibrary) : DL_Process ｜ 版本 (Version) : 1.0.0 ｜ 2026-11-24
 * 兼容性   (Platform)   : CODESYS 3.5+ / TwinCAT 3 / 汇川 InoProShop / 施耐德 Machine Expert
 *                         仅依赖 IEC 61131-3 标准库（TON / R_TRIG / ABS / LIMIT），零厂商私有库
 * 功能描述 (Function)   : 曝气风机间歇循环 + 溶解氧（DO）带控制：DO < fDoLow → eBlowing
 *                         （先开 1 台；若一个 tBlowOn 窗后 DO 仍低于下限则再增开一台，最多
 *                         nBlowerCnt 台）；DO ≥ fDoHigh 且已满足最短曝气 tBlowOn → eResting（全停）；
 *                         eResting 满足最短停曝 tBlowOff 且 DO < fDoLow → 回 eBlowing。
 *                         **迟滞带**：DO ∈ [fDoLow, fDoHigh) 时保持当前相（禁抖，只在两阈值处置位）。
 *                         **仪表失效判据**：DO 采样非有限 → 故障级 eNonFinite；DO 变化量
 *                         |Δ| < 1.0E-6 持续 tDoTimeout（数值完全冻结）→ 故障级 eDoSensorStuck。
 *                         **风机降级**：运行中某台持续无反馈达 3s → 该台置失效标记并停机，
 *                         由台数调节逻辑自动补开备台（信息级 eBlowerSwap，不锁存）；
 *                         无可补备台而需求 > 0 时 → 故障级 eNoBlowerAvail。
 *                         **bStart = FALSE 语义（R191 二选一，本件选「降级为安全值 + 置标志」）**：
 *                         全部风机停、eIdle（曝气风机不得冻结保持）。
 * 接口     (Interface)  : 输入 bEnable / bStart / bReset（上升沿）/ fDoPv / fDoLow / fDoHigh /
 *                         tBlowOn / tBlowOff / tDoTimeout / nBlowerCnt / aBlowerFb[1..3]；
 *                         输出 aBlowerRun[1..3] / nBlowerUsed / eState（E_DL_AbcPhase）/
 *                         eCause（E_DL_AbcCause）/ bError / bValid / tCycleElapsed。
 * 状态迁移表 (State Transition Table)：
 *   ① eIdle → eBlowing：bEnable 且 bStart 且组态闸通过且 fDoPv < fDoLow 且无锁存；
 *      拍 N 进入 / 本拍行为：清失效标记、需求台数置 1、_diCycleMs 清零 / 拍 N+1 转出至 eBlowing。
 *   ② eBlowing → eResting：fDoPv ≥ fDoHigh 且 _bMinOnDone（最短曝气已满足，迟滞上沿）；
 *      拍 N 进入 / 本拍行为：全部风机停、需求台数置 0、_bMinOffDone 复位、_diCycleMs 清零 /
 *      拍 N+1 转出至 eResting。
 *   ③ eBlowing → eBlowing（增台）：tonBlowOn.Q 且 fDoPv 仍 < fDoLow 且需求 < nBlowerCnt；
 *      拍 N 进入（一个曝气窗结束）/ 本拍行为：需求台数 +1、信息级 eBlowerAdded /
 *      拍 N+1 转出（仍在本相，台数调节逻辑补开一台）。
 *   ④ eResting → eBlowing：_bMinOffDone 且 fDoPv < fDoLow（迟滞下沿）；拍 N 进入 /
 *      本拍行为：需求台数置 1、_bMinOnDone 复位、_diCycleMs 清零 / 拍 N+1 转出至 eBlowing。
 *   ⑤ eBlowing → eFault：无可补备台而需求台数 > 0（eNoBlowerAvail）；DO 冻结超时
 *      （eDoSensorStuck）；DO 非有限（eNonFinite）。锁存后由段尾迁移闸迁相（R21）。
 *   ⑥ eFault → eIdle：bReset 上升沿（R_TRIG 判 .Q）且 bEnable = FALSE（R19 穷举出口）；
 *      拍 N 进入 / 本拍行为：清锁存与成因、全部风机停 / 拍 N+1 转出至 eIdle。
 *   ⑦ ELSE（非法枚举值）→ eFault，成因 eIllegalState（R6 兜底）。
 * 边界     (Boundary)   : ① 五个 TON（tonBlowOn / tonBlowOff / tonDoStuck / tonBlowerFb / tonCycle）
 *                            与 R_TRIG 全在 CASE 外无条件调用（R7）；IN 均含 NOT .Q 自复位项（R188）。
 *                         ② 最短曝气 / 最短停曝是**状态量**（_bMinOnDone / _bMinOffDone，由 tonBlowOn /
 *                            tonBlowOff 首个 Q 置位、换相清零），不是单拍标志 —— 避免「Q 早已过去
 *                            而当拍 DO 尚未到上沿」导致最短时间判据被漏掉（禁挂单拍位，R192 类）。
 *                         ③ tonBlowOn.Q 自复位后周期性再触发，故每个 tBlowOn 窗最多增开一台，
 *                            天然的逐级增台节流；增台上限 nBlowerCnt。
 *                         ④ 台数调节：_nRunCnt（实际运行台数）与 _nWant（需求台数）对齐，单拍最多
 *                            补/停一台；补开取最小可用下标，停机取最大下标（后投先停）。
 *                         ⑤ DO 冻结判据的 Δ 用上一拍快照 _fDoPrev（段尾唯一写入），容差 1.0E-6（R4）。
 *                         ⑥ 数组下标安全：_nClamp := LIMIT(1, nBlowerCnt, 3)，全部 FOR 与下标访问
 *                            只用定长 1..3 与 _nClamp（R17 定长数组）。
 *                         ⑦ 零全局耦合（无 GVL / VAR_EXTERNAL / %I / %Q，R1 / R2）。
 * 码表     (Codes)      : 本件不占用全局数字码位（R297 零码位范式）；出口为 BOOL + ENUM，
 *                         enum E_DL_AbcPhase / E_DL_AbcCause 归属本文件（全库唯一属主，R264）。
 *                         信息级（0..9）永不置 bError；故障级（10 起）赋值处与 _bFaultLatch 三行
 *                         成对（R45），锁存回放至 bReset 沿（FB33-1）。
 * 分工声明 (Scope)      : DO 闭环（鼓风机变频 / 阀门开度 PID）归 FB_DL_DoControlLoop 类件；
 *                         曝气池工艺模型与DO预测归高级算法件；本件只做**间歇曝气时序 + 台数分级 +
 *                         DO 迟滞带**，不做连续闭环，也不做鼓风机电机保护。
 * 归属     (Ownership)  : E_DL_AbcPhase / E_DL_AbcCause 归属本文件（全库唯一定义，R264）。
 * 红线自检 (Redline)    : R1 ✓ 零 GVL ｜ R2 ✓ 零 %I/%Q ｜ R3 ✓ 纯 IEC ｜ R4 ✓ 无除法 + 容差比较 +
 *                         非有限双判 ｜ R5 ✓ 逐行同行双语注释 ｜ R6 ✓ 四态 ENUM + CASE + ELSE
 *                         R7 ✓ 全部 TON/R_TRIG 在 CASE 外 ｜ R8/R9 N/A（无 METHOD）｜ R10 ✓ 无构造式
 *                         转换 ｜ R14 ✓ 无 PROPERTY ｜ R15 ✓ 无保留字撞名（aBlowerRun 多字母数组名）
 *                         R17 ✓ 定长 ARRAY[1..3] ｜ R18 ✓ bReset 用 R_TRIG 判 .Q ｜ R19 ✓ eFault
 *                         出口 = bReset 沿 + 撤使能 ｜ R20 ✓ 等待收敛相带超时 ｜ R21 ✓ 锁存与迁相分离。
 * 修订历史 (Revision)   : 2026-11-24  v1.0.0  R79-B 首版
 * 验收向量 (Acceptance) :
 *   V1 fDoLow=2.0、fDoHigh=4.0、tBlowOn=T#30S、tBlowOff=T#60S、nBlowerCnt=2、aBlowerFb 全 TRUE：
 *      fDoPv=1.5 → eBlowing、nBlowerUsed=1、aBlowerRun[1]=TRUE；fDoPv 升至 4.5 且已过 30s →
 *      eResting、nBlowerUsed=0；tBlowOff 到且 fDoPv=1.0 → 回 eBlowing、nBlowerUsed=1。
 *   V2 fDoPv 恒 1.5、nBlowerCnt=3：首个 tBlowOn 窗后 nBlowerUsed=2（eCause=eBlowerAdded），
 *      第二个窗后 nBlowerUsed=3；此后保持 3 台（不再增，信息级 eAllBlowersBusy）。
 *   V3 fDoLow=4.0、fDoHigh=2.0（阈值倒置）→ eState=eFault、eCause=eBadConfig、bError=TRUE、
 *      全部 aBlowerRun=FALSE；bReset 上升沿且 bEnable=FALSE → 回 eIdle、bError=FALSE。
 *   V4 fDoPv 恒为 2.5（|Δ| = 0）持续 tDoTimeout=T#60S → eState=eFault、
 *      eCause=eDoSensorStuck、bError=TRUE。
 *   V5 nBlowerCnt=2、1# 运行中 aBlowerFb[1] 保持 FALSE 超 3s → 1# 停、nBlowerUsed 仍为 1
 *      （2# 补开）、eCause=eBlowerSwap、bError=FALSE（台级降级不锁存）。
 *   V6 nBlowerCnt=1 且该台失效（无备台）→ eState=eFault、eCause=eNoBlowerAvail、bError=TRUE。
 *============================================================================*)

(*-----------------------------------------------------------------------------
 * 枚举: E_DL_AbcPhase（曝气间歇循环相位；eFault 为安全相，仅 bReset 沿迁出）
 *----------------------------------------------------------------------------*)
TYPE E_DL_AbcPhase :
(
    eIdle    := 0,    // 空闲：全部风机停，等启动条件 / Idle: all blowers off, waiting for the start condition
    eBlowing := 10,   // 曝气相：按 DO 逐级开风机 / Blowing: stage blowers up according to the DO
    eResting := 20,   // 停曝相：全部风机停，等最短停曝与 DO 回落 / Resting: all off, waiting for min off time and DO drop
    eFault   := 90    // 故障安全相：锁存成因，全部风机停 / Fault safe phase: latched cause, all blowers off
);
END_TYPE

(*-----------------------------------------------------------------------------
 * 枚举: E_DL_AbcCause（成因码；信息级 = 0..9，故障级 = 10 起）
 *----------------------------------------------------------------------------*)
TYPE E_DL_AbcCause :
(
    eNone            := 0,   // 信息级：无事件 / Info: no event
    eBlowingCode     := 1,   // 信息级：曝气中 / Info: blowing in progress
    eRestingCode     := 2,   // 信息级：停曝中 / Info: resting in progress
    eBlowerAdded     := 3,   // 信息级：低氧未改善，增开一台 / Info: DO still low, one more blower added
    eBlowerSwap      := 4,   // 信息级：台级失效，换备台运行 / Info: one blower failed, standby started instead
    eAllBlowersBusy  := 5,   // 信息级：已达最大台数仍低氧，保持并等工艺 / Info: all blowers running, DO still low
    eBadConfig       := 10,  // 故障级：阈值倒置 / 时间参数越域 / 台数越域 / Fault: inverted thresholds, time or count out of domain
    eNonFinite       := 11,  // 故障级：DO 采样非有限 / Fault: non-finite DO sample
    eDoSensorStuck   := 12,  // 故障级：DO 数值冻结超时（仪表失效）/ Fault: DO frozen beyond the timeout
    eNoBlowerAvail   := 13,  // 故障级：无可补备台而需求台数 > 0 / Fault: demand positive but no blower available
    eIllegalState    := 14   // 故障级：非法状态枚举值 / Fault: illegal state enum value
);
END_TYPE

FUNCTION_BLOCK FB_DL_AerationBlowerCycle
VAR_INPUT
    bEnable      : BOOL := FALSE;             // 使能：FALSE 全部风机停并回 eIdle / Enable, FALSE stops all blowers and returns to idle
    bStart       : BOOL := FALSE;             // 启动（电平）：FALSE 全部风机停 / Start level, FALSE stops all blowers
    bReset       : BOOL := FALSE;             // 复位（上升沿，需同时 bEnable=FALSE）/ Reset rising edge, requires bEnable FALSE
    fDoPv        : LREAL := 0.0;              // 溶解氧实测值 [mg/L] / Measured dissolved oxygen
    fDoLow       : LREAL := 2.0;              // DO 下限（低于即需曝气），域 < fDoHigh [mg/L] / DO low limit, domain < fDoHigh
    fDoHigh      : LREAL := 4.0;              // DO 上限（达此可停曝），域 > fDoLow [mg/L] / DO high limit, domain > fDoLow
    tBlowOn      : TIME := T#30S;             // 最短曝气时长 / 增台窗，域 ≥ 100ms [s] / Minimum blow time and staging window
    tBlowOff     : TIME := T#60S;             // 最短停曝时长，域 ≥ 100ms [s] / Minimum rest time
    tDoTimeout   : TIME := T#60S;             // DO 冻结判失效超时，域 100ms..1h [s] / DO frozen-to-fail timeout
    nBlowerCnt   : INT := 2;                  // 装机风机台数，有效域 1..3 [台] / Installed blower count, valid domain 1..3
    aBlowerFb    : ARRAY[1..3] OF BOOL;       // 各风机运行反馈（TRUE = 在转）[#] / Per-blower running feedback
END_VAR
VAR_OUTPUT
    aBlowerRun   : ARRAY[1..3] OF BOOL;       // 各风机启动命令（内部状态映射，段 8 单点出口）[#] / Per-blower run command mapped at the tail
    nBlowerUsed  : INT := 0;                  // 当前运行风机台数 [台] / Number of running blowers
    eState       : E_DL_AbcPhase;             // 状态出口（段尾单点映射）[-] / State outlet mapped at the tail
    eCause       : E_DL_AbcCause;             // 成因码出口（故障期锁存回放）[-] / Cause code outlet
    bError       : BOOL;                      // 故障锁存标志 [-] / Fault latch flag
    bValid       : BOOL;                      // 循环有效回执（曝气/停曝相且无锁存）[-] / Cycle validity receipt
    tCycleElapsed : TIME := T#0S;             // 当前相驻留时长 [s] / Dwell time of the current phase
END_VAR
VAR
    _eState       : E_DL_AbcPhase := E_DL_AbcPhase.eIdle;   // 内部相位（CASE 唯一写入目标）[-] / Internal phase
    _bFaultLatch  : BOOL := FALSE;                          // 故障锁存位（仅 bReset 沿清除）[-] / Fault latch bit
    _eCauseLatch  : E_DL_AbcCause := E_DL_AbcCause.eNone;    // 锁存成因码（FB33-1 锁存回放）[-] / Latched cause code
    _eCauseTmp    : E_DL_AbcCause := E_DL_AbcCause.eNone;    // 本拍首因中间量（段 7 组态闸用）[-] / First cause of this scan
    _bCfgOk       : BOOL := TRUE;                           // 组态与入参闸通过标志 [-] / Configuration gate flag
    _bResetPulse  : BOOL := FALSE;                          // bReset 上升沿快照（R18）[-] / bReset rising-edge snapshot
    _nClamp       : INT := 1;                               // 装机台数钳位值 1..3 [台] / Clamped installed blower count
    _nIdx         : INT := 1;                               // 遍历下标（FOR 专用）[台] / Loop index for FOR statements
    _nPick        : INT := 0;                               // 本拍选中风机下标，0 = 未选中 [台] / Blower index picked in this scan
    _nWant        : INT := 0;                               // 需求运行台数 [台] / Required number of running blowers
    _nRunCnt      : INT := 0;                               // 实际运行台数（含未确认反馈者）[台] / Actual running blower count
    _nFbSuspect   : INT := 0;                               // 无反馈嫌疑风机下标，0 = 无 [台] / Suspect blower index without feedback
    _aBlowerRun   : ARRAY[1..3] OF BOOL;                    // 内部启动命令状态数组 [#] / Internal run-command state array
    _aBlowerBad   : ARRAY[1..3] OF BOOL;                    // 内部台级失效标记（换备台用，eIdle 清除）[#] / Internal per-blower failure flags
    _bMinOnDone   : BOOL := FALSE;                          // 最短曝气已满足（状态量，非单拍位）[-] / Min blow time satisfied, a state not a pulse
    _bMinOffDone  : BOOL := FALSE;                          // 最短停曝已满足（状态量，非单拍位）[-] / Min rest time satisfied, a state not a pulse
    _fDoPrev      : LREAL := 0.0;                           // 上一拍 DO 快照（冻结判据用，段尾唯一写入）[mg/L] / DO snapshot of the last scan
    _bDoMoving    : BOOL := FALSE;                          // DO 本拍有变化标志 [-] / DO changed in this scan
    _diCycleMs    : DINT := 0;                              // 当前相驻留毫秒累加 [ms] / Accumulated dwell milliseconds
    rtReset       : R_TRIG;                                 // bReset 边沿实例（段 4 无条件调用，R18）/ bReset edge instance called unconditionally
    tonBlowOn     : TON;                                    // 最短曝气 / 增台窗定时器（段 4 无条件调用）/ Min blow and staging window timer
    tonBlowOff    : TON;                                    // 最短停曝定时器（段 4 无条件调用）/ Min rest timer called unconditionally
    tonDoStuck    : TON;                                    // DO 冻结持续判（段 4 无条件调用）/ DO frozen persistence timer
    tonBlowerFb   : TON;                                    // 单台无反馈持续判（段 4 无条件调用）/ Per-blower feedback loss timer
    tonCycle      : TON;                                    // 相驻留时长采样节拍（段 4 无条件调用）/ Dwell-time sampling tick
END_VAR
VAR CONSTANT
    DL_ABC_ZERO      : LREAL := 0.0;             // 浮点零基准 [-] / Float zero base
    DL_ABC_EPS       : LREAL := 1.0E-6;          // DO 变化量容差（冻结判据）[mg/L] / DO change tolerance for the freeze check
    DL_ABC_BLOWER_MAX : INT := 3;                // 风机台数上限（数组定长）[台] / Upper bound of blowers, fixed array size
    DL_ABC_ONE       : INT := 1;                 // 台数起始值 [台] / Count start value
    DL_ABC_FB_WIN    : TIME := T#3S;             // 单台无反馈持续窗 [s] / Per-blower feedback loss window
    DL_ABC_T_MIN     : TIME := T#100MS;          // 时间参数下限 [s] / Lower bound of the time parameters
    DL_ABC_T_MAX     : TIME := T#1H;             // 时间参数上限 [s] / Upper bound of the time parameters
    DL_ABC_DT        : TIME := T#100MS;          // 驻留时长采样节拍 [s] / Dwell-time sampling tick
    DL_ABC_DT_MS     : DINT := 100;              // 采样节拍毫秒数 [ms] / Sampling tick in milliseconds
    DL_ABC_MS_ZERO   : DINT := 0;                // 毫秒零基准 [-] / Millisecond zero base
END_VAR

(* —— 段 1：中间量预置（不清锁存 / 数组状态 / 驻留累加，FB32-1） —— *)
_bCfgOk    := TRUE;                                    // 组态闸标志复位 / Configuration flag reset
_eCauseTmp := E_DL_AbcCause.eNone;                      // 当拍首因复位 / Scan cause reset
_nPick     := 0;                                       // 选中下标复位 / Picked index reset
_bDoMoving := FALSE;                                   // DO 变化标志复位 / DO change flag reset

(* —— 段 2：台数钳位与 DO 变化判据（浮点容差比较，R4） —— *)
_nClamp := LIMIT(DL_ABC_ONE, nBlowerCnt, DL_ABC_BLOWER_MAX);            // 台数钳位 1..3 / Clamp the blower count
IF ABS(fDoPv - _fDoPrev) >= DL_ABC_EPS THEN
    _bDoMoving := TRUE;                                                 // Δ 达容差：DO 在变化 / Delta above tolerance: DO is moving
ELSE
    _bDoMoving := FALSE;                                                // Δ 小于容差：本拍视作冻结 / Delta below tolerance: frozen this scan
END_IF

(* —— 段 3：组态与入参域闸（阈值倒置 / 时间越域 / 台数越域 / 非有限） —— *)
IF (fDoPv <> fDoPv) OR ((fDoPv - fDoPv) <> DL_ABC_ZERO)
    OR (fDoLow <> fDoLow) OR ((fDoLow - fDoLow) <> DL_ABC_ZERO)
    OR (fDoHigh <> fDoHigh) OR ((fDoHigh - fDoHigh) <> DL_ABC_ZERO) THEN
    _bCfgOk    := FALSE;                               // 入参非有限 / Non-finite input
    _eCauseTmp := E_DL_AbcCause.eNonFinite;            // 故障级：非有限入参 / Fault: non-finite input
END_IF
IF _bCfgOk THEN
    IF fDoLow >= fDoHigh THEN
        _bCfgOk    := FALSE;                           // 阈值倒置（或无迟滞带）/ Inverted thresholds, no hysteresis band
        _eCauseTmp := E_DL_AbcCause.eBadConfig;        // 故障级：组态非法 / Fault: bad configuration
    ELSIF (nBlowerCnt < DL_ABC_ONE) OR (nBlowerCnt > DL_ABC_BLOWER_MAX) THEN
        _bCfgOk    := FALSE;                           // 装机台数越域 / Blower count out of domain
        _eCauseTmp := E_DL_AbcCause.eBadConfig;        // 故障级：组态非法 / Fault: bad configuration
    ELSIF (tBlowOn < DL_ABC_T_MIN) OR (tBlowOn > DL_ABC_T_MAX) THEN
        _bCfgOk    := FALSE;                           // 最短曝气越域 / Min blow time out of domain
        _eCauseTmp := E_DL_AbcCause.eBadConfig;        // 故障级：组态非法 / Fault: bad configuration
    ELSIF (tBlowOff < DL_ABC_T_MIN) OR (tBlowOff > DL_ABC_T_MAX) THEN
        _bCfgOk    := FALSE;                           // 最短停曝越域 / Min rest time out of domain
        _eCauseTmp := E_DL_AbcCause.eBadConfig;        // 故障级：组态非法 / Fault: bad configuration
    ELSIF (tDoTimeout < DL_ABC_T_MIN) OR (tDoTimeout > DL_ABC_T_MAX) THEN
        _bCfgOk    := FALSE;                           // DO 冻结超时越域 / DO freeze timeout out of domain
        _eCauseTmp := E_DL_AbcCause.eBadConfig;        // 故障级：组态非法 / Fault: bad configuration
    END_IF
END_IF

(* —— 段 4：边沿与定时器（CASE 外无条件调用，R7；IN 均含 NOT .Q 自复位，R188） —— *)
rtReset(CLK := bReset);                                // bReset 边沿无条件刷新（R18）/ bReset edge refreshed unconditionally
_bResetPulse := rtReset.Q;                             // 边沿快照 / Edge snapshot
tonBlowOn(IN := (_eState = E_DL_AbcPhase.eBlowing) AND (NOT tonBlowOn.Q) AND (NOT _bFaultLatch),
          PT := tBlowOn);                              // 最短曝气 / 增台窗（自复位后周期性再触发）/ Min blow and staging window
tonBlowOff(IN := (_eState = E_DL_AbcPhase.eResting) AND (NOT tonBlowOff.Q) AND (NOT _bFaultLatch),
           PT := tBlowOff);                            // 最短停曝（自复位后周期性再触发）/ Min rest window
tonCycle(IN := ((_eState = E_DL_AbcPhase.eBlowing) OR (_eState = E_DL_AbcPhase.eResting))
              AND (NOT tonCycle.Q) AND (NOT _bFaultLatch),
         PT := DL_ABC_DT);                             // 相驻留时长采样节拍 / Dwell-time sampling tick
IF tonCycle.Q THEN
    _diCycleMs := _diCycleMs + DL_ABC_DT_MS;           // 驻留毫秒累加 / Accumulate dwell milliseconds
END_IF
(* 无反馈嫌疑台：取最小下标的「已命令但无反馈」风机（用上一拍状态，一拍延迟） *)
_nFbSuspect := 0;                                      // 嫌疑下标复位 / Suspect index reset
FOR _nIdx := 1 TO DL_ABC_BLOWER_MAX DO
    IF (_nFbSuspect = 0) AND _aBlowerRun[_nIdx] AND (NOT aBlowerFb[_nIdx]) THEN
        _nFbSuspect := _nIdx;                          // 记录首个无反馈风机 / Record the first blower without feedback
    END_IF
END_FOR
tonBlowerFb(IN := (_nFbSuspect > 0) AND (NOT tonBlowerFb.Q) AND (NOT _bFaultLatch),
            PT := DL_ABC_FB_WIN);                      // 单台无反馈持续判 / Per-blower feedback loss persistence
tonDoStuck(IN := bEnable AND bStart AND (NOT _bDoMoving)
                AND (NOT tonDoStuck.Q) AND (NOT _bFaultLatch),
           PT := tDoTimeout);                          // DO 冻结持续判（仪表失效）/ DO frozen persistence check

(* —— 段 5：状态机主体（唯一相位写入点；故障只置锁存，迁相由段 7 统一执行） —— *)
CASE _eState OF
    E_DL_AbcPhase.eIdle :
        FOR _nIdx := 1 TO DL_ABC_BLOWER_MAX DO
            _aBlowerRun[_nIdx] := FALSE;               // 空闲：命令全撤 / Idle: commands withdrawn
            _aBlowerBad[_nIdx] := FALSE;               // 空闲：台级失效标记清除 / Idle: failure flags cleared
        END_FOR
        _nWant      := 0;                              // 空闲：需求台数 0 / Idle: demand zero
        _nRunCnt    := 0;                              // 空闲：运行台数 0 / Idle: run count zero
        _bMinOnDone := FALSE;                          // 空闲：最短曝气状态复位 / Idle: min-blow state cleared
        _bMinOffDone := FALSE;                         // 空闲：最短停曝状态复位 / Idle: min-rest state cleared
        _diCycleMs  := DL_ABC_MS_ZERO;                 // 空闲：驻留累计清零 / Idle: dwell accumulator cleared
        IF bEnable AND bStart AND _bCfgOk AND (fDoPv < fDoLow) AND (NOT _bFaultLatch) THEN
            _nWant      := DL_ABC_ONE;                 // 迁移①：先开 1 台 / Start with one blower
            _bMinOnDone := FALSE;                      // 最短曝气状态复位 / Min-blow state cleared
            _bMinOffDone := FALSE;                     // 最短停曝状态复位 / Min-rest state cleared
            _diCycleMs  := DL_ABC_MS_ZERO;             // 驻留累计清零 / Dwell accumulator cleared
            eCause      := E_DL_AbcCause.eBlowingCode; // 信息级：开始曝气 / Info: blowing started
            _eState     := E_DL_AbcPhase.eBlowing;     // 进入曝气相 / Move to blowing
        END_IF

    E_DL_AbcPhase.eBlowing :
        IF (NOT bEnable) OR (NOT bStart) THEN
            FOR _nIdx := 1 TO DL_ABC_BLOWER_MAX DO
                _aBlowerRun[_nIdx] := FALSE;           // 失能：命令全撤 / Disabled: all commands withdrawn
            END_FOR
            _nWant      := 0;                          // 需求台数 0 / Demand zero
            _nRunCnt    := 0;                          // 运行台数 0 / Run count zero
            _diCycleMs  := DL_ABC_MS_ZERO;             // 驻留累计清零 / Dwell accumulator cleared
            eCause      := E_DL_AbcCause.eNone;        // 信息级：无事件 / Info: no event
            _eState     := E_DL_AbcPhase.eIdle;        // 回空闲相 / Back to idle
        ELSE
            (* 最长曝气窗到：置最短曝气满足状态量（非单拍位）/ 低氧未改善则逐级增台 *)
            IF tonBlowOn.Q THEN
                _bMinOnDone := TRUE;                   // 最短曝气已满足（状态量）/ Min blow satisfied as a state
                IF fDoPv < fDoLow THEN
                    IF _nWant < _nClamp THEN
                        _nWant := _nWant + DL_ABC_ONE; // 迁移③：低氧未改善，需求 +1 / DO still low: demand plus one
                        eCause := E_DL_AbcCause.eBlowerAdded;   // 信息级：增开一台 / Info: one blower added
                    ELSE
                        eCause := E_DL_AbcCause.eAllBlowersBusy; // 信息级：已达最大台数 / Info: all blowers already running
                    END_IF
                END_IF
            END_IF
            (* 台级反馈丢失降级：嫌疑台置失效、停机，随后由台数调节补开备台 *)
            IF tonBlowerFb.Q AND (_nFbSuspect > 0) THEN
                IF (_nFbSuspect >= DL_ABC_ONE) AND (_nFbSuspect <= DL_ABC_BLOWER_MAX) THEN
                    _aBlowerBad[_nFbSuspect] := TRUE;  // 该台置失效标记 / Mark this blower as failed
                    IF _aBlowerRun[_nFbSuspect] THEN
                        _aBlowerRun[_nFbSuspect] := FALSE;   // 撤该台命令 / Withdraw this command
                        IF _nRunCnt > 0 THEN
                            _nRunCnt := _nRunCnt - DL_ABC_ONE; // 运行台数回退 / Roll the run count back
                        END_IF
                    END_IF
                    eCause := E_DL_AbcCause.eBlowerSwap;     // 信息级：台级失效换备台 / Info: failed blower swapped out
                END_IF
            END_IF
            (* 台数调节：需求与实际对齐，单拍最多补/停一台 *)
            IF _nRunCnt < _nWant THEN
                _nPick := 0;                           // 补开候选复位 / Candidate reset
                FOR _nIdx := 1 TO _nClamp DO
                    IF (_nPick = 0) AND (NOT _aBlowerRun[_nIdx]) AND (NOT _aBlowerBad[_nIdx]) THEN
                        _nPick := _nIdx;               // 取最小可用下标（未运行且未失效）/ Lowest available blower
                    END_IF
                END_FOR
                IF _nPick > 0 THEN
                    _aBlowerRun[_nPick] := TRUE;       // 补开一台 / Start one blower
                    _nRunCnt := _nRunCnt + DL_ABC_ONE; // 运行台数 +1 / Increment the run count
                ELSE
                    IF NOT _bFaultLatch THEN
                        _eCauseLatch := E_DL_AbcCause.eNoBlowerAvail;   // 故障级：无可补备台 / Fault: no blower available
                        _bFaultLatch := TRUE;                           // 置故障锁存（迁相由段 7，R21）/ Latch the fault
                    END_IF
                END_IF
            ELSIF _nRunCnt > _nWant THEN
                _nPick := 0;                           // 停机候选复位 / Stop candidate reset
                FOR _nIdx := 1 TO _nClamp DO
                    IF _aBlowerRun[_nIdx] THEN
                        _nPick := _nIdx;               // 取最大下标（后投先停）/ Highest index, last started first stopped
                    END_IF
                END_FOR
                IF _nPick > 0 THEN
                    _aBlowerRun[_nPick] := FALSE;      // 停一台 / Stop one blower
                    _nRunCnt := _nRunCnt - DL_ABC_ONE; // 运行台数 -1 / Decrement the run count
                END_IF
            END_IF
            (* 停曝判据：DO 达上沿且最短曝气已满足（迟滞上沿，R4 大小判据） *)
            IF (fDoPv >= fDoHigh) AND _bMinOnDone THEN
                FOR _nIdx := 1 TO DL_ABC_BLOWER_MAX DO
                    _aBlowerRun[_nIdx] := FALSE;       // 迁移②：全部风机停 / All blowers stopped
                END_FOR
                _nWant      := 0;                      // 需求台数 0 / Demand zero
                _nRunCnt    := 0;                      // 运行台数 0 / Run count zero
                _bMinOffDone := FALSE;                 // 最短停曝状态复位 / Min-rest state cleared
                _diCycleMs  := DL_ABC_MS_ZERO;         // 驻留累计清零 / Dwell accumulator cleared
                eCause      := E_DL_AbcCause.eRestingCode;   // 信息级：进入停曝 / Info: resting started
                _eState     := E_DL_AbcPhase.eResting; // 进入停曝相 / Move to resting
            ELSE
                IF eCause = E_DL_AbcCause.eNone THEN
                    eCause := E_DL_AbcCause.eBlowingCode;    // 信息级：曝气中 / Info: blowing in progress
                END_IF
            END_IF
        END_IF

    E_DL_AbcPhase.eResting :
        FOR _nIdx := 1 TO DL_ABC_BLOWER_MAX DO
            _aBlowerRun[_nIdx] := FALSE;               // 停曝相：命令全撤 / Resting: all commands withdrawn
        END_FOR
        _nWant   := 0;                                 // 需求台数 0 / Demand zero
        _nRunCnt := 0;                                 // 运行台数 0 / Run count zero
        IF (NOT bEnable) OR (NOT bStart) THEN
            _diCycleMs := DL_ABC_MS_ZERO;              // 驻留累计清零 / Dwell accumulator cleared
            eCause     := E_DL_AbcCause.eNone;         // 信息级：无事件 / Info: no event
            _eState    := E_DL_AbcPhase.eIdle;         // 回空闲相 / Back to idle
        ELSE
            IF tonBlowOff.Q THEN
                _bMinOffDone := TRUE;                  // 最短停曝已满足（状态量）/ Min rest satisfied as a state
            END_IF
            IF _bMinOffDone AND (fDoPv < fDoLow) THEN
                _nWant      := DL_ABC_ONE;             // 迁移④：下限已触发，先开 1 台 / Low limit reached: start with one
                _bMinOnDone := FALSE;                  // 最短曝气状态复位 / Min-blow state cleared
                _diCycleMs  := DL_ABC_MS_ZERO;         // 驻留累计清零 / Dwell accumulator cleared
                eCause      := E_DL_AbcCause.eBlowingCode;   // 信息级：恢复曝气 / Info: blowing resumed
                _eState     := E_DL_AbcPhase.eBlowing; // 进入曝气相 / Move to blowing
            ELSE
                eCause := E_DL_AbcCause.eRestingCode;  // 信息级：停曝中（迟滞带内保持）/ Info: resting in progress
            END_IF
        END_IF

    E_DL_AbcPhase.eFault :
        FOR _nIdx := 1 TO DL_ABC_BLOWER_MAX DO
            _aBlowerRun[_nIdx] := FALSE;               // 故障相：命令全撤（安全侧）/ Fault phase: all commands withdrawn
        END_FOR
        _nWant     := 0;                               // 需求台数 0 / Demand zero
        _nRunCnt   := 0;                               // 运行台数 0 / Run count zero
        _diCycleMs := DL_ABC_MS_ZERO;                  // 驻留累计清零 / Dwell accumulator cleared
        IF _bResetPulse AND (NOT bEnable) THEN
            _bFaultLatch := FALSE;                     // 迁移⑥：清故障锁存 / Clear the fault latch
            _eCauseLatch := E_DL_AbcCause.eNone;       // 清锁存成因 / Clear the latched cause
            eCause       := E_DL_AbcCause.eNone;       // 出口同步归零 / Outlet follows
            _bMinOnDone  := FALSE;                     // 最短曝气状态复位 / Min-blow state cleared
            _bMinOffDone := FALSE;                     // 最短停曝状态复位 / Min-rest state cleared
            _eState      := E_DL_AbcPhase.eIdle;       // 回空闲相 / Back to idle
        END_IF

ELSE
    (* 迁移⑦：非法枚举兜底（R6） *)
    IF NOT _bFaultLatch THEN
        _eCauseLatch := E_DL_AbcCause.eIllegalState;   // 故障级：非法状态 / Fault: illegal state
        _bFaultLatch := TRUE;                          // 置故障锁存 / Latch the fault
    END_IF
END_CASE

(* —— 段 6：DO 冻结超时（仪表失效）的锁存（锁存与迁相分离，R21） —— *)
IF tonDoStuck.Q AND (NOT _bFaultLatch) THEN
    _eCauseLatch := E_DL_AbcCause.eDoSensorStuck;      // 故障级：DO 数值冻结 / Fault: DO value frozen
    _bFaultLatch := TRUE;                              // 置故障锁存 / Latch the fault
END_IF

(* —— 段 7：组态闸失败处理 + 段尾故障迁移闸 + 故障相动作全撤（FB50-1④） —— *)
IF (NOT _bCfgOk) AND (NOT _bFaultLatch) THEN
    _eCauseLatch := _eCauseTmp;                        // 锁存首因（组态闸）/ Latch the configuration cause
    _bFaultLatch := TRUE;                              // 置故障锁存 / Latch the fault
END_IF
IF _bFaultLatch AND (_eState <> E_DL_AbcPhase.eFault) THEN
    _eState := E_DL_AbcPhase.eFault;                   // 锁存即迁相 / Latch forces the fault phase
END_IF
IF _eState = E_DL_AbcPhase.eFault THEN
    FOR _nIdx := 1 TO DL_ABC_BLOWER_MAX DO
        _aBlowerRun[_nIdx] := FALSE;                   // 故障相命令全撤（含同拍迁入）/ All commands withdrawn in fault
    END_FOR
    _nWant   := 0;                                     // 需求台数 0 / Demand zero
    _nRunCnt := 0;                                     // 运行台数 0 / Run count zero
END_IF

(* —— 段 8：统一出口（状态映射 + 台数映射 + 驻留换算 + 锁存回放） —— *)
eState := _eState;                                     // 相位映射 / Phase mapping
FOR _nIdx := 1 TO DL_ABC_BLOWER_MAX DO
    aBlowerRun[_nIdx] := _aBlowerRun[_nIdx];           // 启动命令映射 / Run command mapping
END_FOR
nBlowerUsed   := _nRunCnt;                             // 运行台数出口 / Running count outlet
tCycleElapsed := DINT_TO_TIME(_diCycleMs);             // 驻留毫秒 → TIME（标准转换，R10）/ Dwell milliseconds to TIME
bError := _bFaultLatch;                                // 故障标志取锁存位 / Fault flag from the latch
IF _bFaultLatch THEN
    eCause := _eCauseLatch;                            // 故障期回放锁存码（FB33-1）/ Replay the latched code
END_IF
bValid := ((_eState = E_DL_AbcPhase.eBlowing) OR (_eState = E_DL_AbcPhase.eResting))
          AND (NOT _bFaultLatch);                      // 曝气/停曝相且无锁存时有效 / Valid while blowing or resting without a latch
_fDoPrev := fDoPv;                                     // DO 快照更新（唯一写入点，冻结判据用）/ DO snapshot, single write point
END_FUNCTION_BLOCK
